(* IEC 61131-3 sources: volt/packages/volt-lsp-iec/test-corpus/pro2193/Device/Plc Logic/Application/09 Misc/Library Manager/L_TT1P_TechnologyModules, 514 files *)

(* ---- _SCAP_TM_BASICMOTIONBASE.dut ---- *)
TYPE _SCAP_TM_BASICMOTIONBASE :
STRUCT
END_STRUCT
END_TYPE

(* ---- _SCAP_TM_BASICMOTIONHIGH.dut ---- *)
TYPE _SCAP_TM_BASICMOTIONHIGH :
STRUCT
END_STRUCT
END_TYPE

(* ---- _SCAP_TM_BASICMOTIONSTATE.dut ---- *)
TYPE _SCAP_TM_BASICMOTIONSTATE :
STRUCT
END_STRUCT
END_TYPE

(* ---- _SCAP_TM_CROSSCUTTERBASE.dut ---- *)
TYPE _SCAP_TM_CROSSCUTTERBASE :
STRUCT
	AP01_XENDOFPROFILEWINDOWSIZE : BOOL;
	AP01_LRENDOFPROFILEWINDOWSIZE : LREAL := 0;
	AP02_XOVERSPEEDUPPERLIMIT : BOOL;
	AP02_LROVERSPEEDUPPERLIMIT : LREAL := 2;
	AP07_XSETOFFSETSLAVE : BOOL;
	AP07_LRSETOFFSETSLAVE : LREAL;
	AP08_XOFFSETSLAVEPAR : BOOL;
	AP08_LROFFSETSLAVEVEL : LREAL;
	AP08_LROFFSETSLAVEACC : LREAL;
	AP08_LROFFSETSLAVEDEC : LREAL;
	AP08_LROFFSETSLAVEJERK : LREAL;
	AP09_XSETVALUEMODE : BOOL;
	AP09_ESETVALUEMODE : L_MC1P_SetValueMode := L_MC1P_SetValueMode.PosVelAcc;
END_STRUCT
END_TYPE

(* ---- _SCAP_TM_CROSSCUTTERHIGH.dut ---- *)
TYPE _SCAP_TM_CROSSCUTTERHIGH :
STRUCT
END_STRUCT
END_TYPE

(* ---- _SCAP_TM_CROSSCUTTERSTATE.dut ---- *)
TYPE _SCAP_TM_CROSSCUTTERSTATE :
STRUCT
	AP03_XTPAXISDELAYCYCLE : BOOL;
	AP03_LRTPAXISDELAYCYCLE : LREAL;
	AP04_XTPAXISCOMPFACTOR : BOOL;
	AP04_LRTPAXISCOMPFACTOR : LREAL;
	AP05_XUPPERCORRPOS : BOOL;
	AP05_LRUPPERCORRPOS : LREAL;
	AP06_XLOWERCORRPOS : BOOL;
	AP06_LRLOWERCORRPOS : LREAL;
	AP10_XCUTTINGANGLESTOPCAM : BOOL;
	AP10_LRCUTTINGANGLESTOPCAM : LREAL := 10;
	AP11_XSETCUTLENGTHINPRODUCT : BOOL;
END_STRUCT
END_TYPE

(* ---- _SCAP_TM_ELECTRICALSHAFTPOSBASE.dut ---- *)
TYPE _SCAP_TM_ELECTRICALSHAFTPOSBASE :
STRUCT
	AP01_XLOADGEARBOXPOSOUT : BOOL;
	AP01_LRLOADGEARBOXPOSOUT : LREAL;
END_STRUCT
END_TYPE

(* ---- _SCAP_TM_ELECTRICALSHAFTPOSHIGH.dut ---- *)
TYPE _SCAP_TM_ELECTRICALSHAFTPOSHIGH :
STRUCT
	AP05_XLOADOFFSETSYNC : BOOL;
	AP05_LRLOADOFFSETSYNC : LREAL;
END_STRUCT
END_TYPE

(* ---- _SCAP_TM_ELECTRICALSHAFTPOSSTATE.dut ---- *)
TYPE _SCAP_TM_ELECTRICALSHAFTPOSSTATE :
STRUCT
	AP02_XLOADTRIMOFFSET : BOOL;
	AP02_LRLOADTRIMOFFSET : LREAL;
END_STRUCT
END_TYPE

(* ---- _SCAP_TM_ELECTRICALSHAFTVELBASE.dut ---- *)
TYPE _SCAP_TM_ELECTRICALSHAFTVELBASE :
STRUCT
	AP01_XCOUPLINGX : BOOL;
	AP01_LRCOUPLINGX : LREAL := 1.0;
	AP02_XCOUPLINGY : BOOL;
	AP02_LRCOUPLINGY : LREAL := 1.0;
END_STRUCT
END_TYPE

(* ---- _SCAP_TM_ELECTRICALSHAFTVELHIGH.dut ---- *)
TYPE _SCAP_TM_ELECTRICALSHAFTVELHIGH :
STRUCT
END_STRUCT
END_TYPE

(* ---- _SCAP_TM_ELECTRICALSHAFTVELSTATE.dut ---- *)
TYPE _SCAP_TM_ELECTRICALSHAFTVELSTATE :
STRUCT
END_STRUCT
END_TYPE

(* ---- _SCAP_TM_FLEXCAMBASE.dut ---- *)
TYPE _SCAP_TM_FLEXCAMBASE :
STRUCT
	AP01_XENDOFPROFILEWINDOWSIZE : BOOL;
	AP01_LRENDOFPROFILEWINDOWSIZE : LREAL := 0;
	AP02_XSETVALUEMODE : BOOL;
	AP02_ESETVALUEMODE : L_MC1P_SetValueMode := L_MC1P_SetValueMode.PosVelAcc;
END_STRUCT
END_TYPE

(* ---- _SCAP_TM_FLEXCAMHIGH.dut ---- *)
TYPE _SCAP_TM_FLEXCAMHIGH :
STRUCT
END_STRUCT
END_TYPE

(* ---- _SCAP_TM_FLEXCAMSTATE.dut ---- *)
TYPE _SCAP_TM_FLEXCAMSTATE :
STRUCT
END_STRUCT
END_TYPE

(* ---- _SCAP_TM_FLYINGSAWBASE.dut ---- *)
TYPE _SCAP_TM_FLYINGSAWBASE :
STRUCT
	AP01_XLOADTOTALCUTTINGLENGTH : BOOL;
	AP01_LRLOADTOTALCUTTINGLENGTH : LREAL;
	AP02_XLOADTARGETPOS : BOOL;
	AP02_LRLOADTARGETPOS : LREAL;
END_STRUCT
END_TYPE

(* ---- _SCAP_TM_FLYINGSAWHIGH.dut ---- *)
TYPE _SCAP_TM_FLYINGSAWHIGH :
STRUCT
	AP02_XLOADTRIMOFFSET : BOOL;
	AP02_LRLOADTRIMOFFSET : LREAL;
END_STRUCT
END_TYPE

(* ---- _SCAP_TM_FLYINGSAWSTATE.dut ---- *)
TYPE _SCAP_TM_FLYINGSAWSTATE :
STRUCT
	AP03_XRANGEOFTOLERANCE : BOOL;
	AP03_LRRANGEOFTOLERANCE : LREAL;
	AP04_XMARKDETECTERRCOMP : BOOL;
	AP04_LRMARKDETECTERRCOMP : LREAL;
	AP05_XTASKCYCLEDELAY : BOOL;
	AP05_BYTASKCYCLEDELAY : BYTE;
END_STRUCT
END_TYPE

(* ---- _SCAP_TM_MOTIONCONTROL.dut ---- *)
TYPE _SCAP_TM_MOTIONCONTROL :
STRUCT
END_STRUCT
END_TYPE

(* ---- _SCAP_TM_PICKANDPLACEBASE.dut ---- *)
TYPE _SCAP_TM_PICKANDPLACEBASE :
STRUCT
	AP01_XCALCPROFILEMOVEPATH : BOOL := TRUE;
END_STRUCT
END_TYPE

(* ---- _SCAP_TM_PICKANDPLACEHIGH.dut ---- *)
TYPE _SCAP_TM_PICKANDPLACEHIGH :
STRUCT
END_STRUCT
END_TYPE

(* ---- _SCAP_TM_PICKANDPLACESTATE.dut ---- *)
TYPE _SCAP_TM_PICKANDPLACESTATE :
STRUCT
	AP02_EBUFFERMODEBLENDING : MC_BUFFER_MODE := MC_BUFFER_MODE.mcBlendingLow;
END_STRUCT
END_TYPE

(* ---- _SCAP_TM_REGISTERCONTROLBASE.dut ---- *)
TYPE _SCAP_TM_REGISTERCONTROLBASE :
STRUCT
	AP03_XTPAXISDELAYCYCLE : BOOL;
	AP03_LRTPAXISDELAYCYCLE : LREAL;
	AP04_XTPAXISCOMPFACTOR : BOOL;
	AP04_LRTPAXISCOMPFACTOR : LREAL;
	AP06_XCORRECTIONONMASTERPOS : BOOL;
	AP07_XLOADSENSORPOS : BOOL;
	AP07_LRLOADSENSORPOS : LREAL;
END_STRUCT
END_TYPE

(* ---- _SCAP_TM_REGISTERCONTROLHIGH.dut ---- *)
TYPE _SCAP_TM_REGISTERCONTROLHIGH :
STRUCT
END_STRUCT
END_TYPE

(* ---- _SCAP_TM_REGISTERCONTROLSTATE.dut ---- *)
TYPE _SCAP_TM_REGISTERCONTROLSTATE :
STRUCT
END_STRUCT
END_TYPE

(* ---- _SCAP_TM_SMARTTRACKBASE.dut ---- *)
TYPE _SCAP_TM_SMARTTRACKBASE :
STRUCT
END_STRUCT
END_TYPE

(* ---- _SCAP_TM_SMARTTRACKHIGH.dut ---- *)
TYPE _SCAP_TM_SMARTTRACKHIGH :
STRUCT
END_STRUCT
END_TYPE

(* ---- _SCAP_TM_SMARTTRACKSTATE.dut ---- *)
TYPE _SCAP_TM_SMARTTRACKSTATE :
STRUCT
	AP_XALLTRACKCORRCAM : BOOL;
	AP_ASCALLTRACKCORRCAM : ARRAY [0..4] OF L_MC2P_XYVA := [STRUCT(eLawOfMotion := L_MC2P_LawOfMotion.Poly5, lrX := 0, lrY := 0, lrYs := 0, lrYss := 0), STRUCT(eLawOfMotion := L_MC2P_LawOfMotion.StraightLine, lrX := 0.179999992251396, lrY := 0.1, lrYs := 1.25000011525118, lrYss := 0), STRUCT(eLawOfMotion := L_MC2P_LawOfMotion.Poly5, lrX := 0.819999933242798, lrY := 0.9, lrYs := 1.25000011525118, lrYss := 0), STRUCT(eLawOfMotion := L_MC2P_LawOfMotion.Poly5, lrX := 1.0, lrY := 1.0, lrYs := 0, lrYss := 0)];
END_STRUCT
END_TYPE

(* ---- _SCAP_TM_STACKERCRANEAXISCONTROLBASE.dut ---- *)
TYPE _SCAP_TM_STACKERCRANEAXISCONTROLBASE :
STRUCT
	AP01_XSETCONTROLLERMODE : BOOL;
	AP01_ECONTROLMODE : L_MC1P_ControlModeSet;
	AP03_XOSCCOMPPOSSCALED : BOOL;
	AP03_LROSCCOMPPOSSCALED : LREAL;
	AP04_XOSCCOMPLOADSCALED : BOOL;
	AP04_LROSCCOMPLOADSCALED : LREAL;
	AP05_EOSCCOMPEXECUTIONINDEX : WORD := 1;
	AP06_XOSCCOMPIGNOREFILTERONSTOP : BOOL := FALSE;
	AP07_XOSCCOMPMANIPULATETROQUE : BOOL := FALSE;
	AP08_XOSCCOMPAMPRATIO : BOOL;
	AP08_LROSCCOMPAMPRATIO : LREAL;
	AP09_XOSCCOMPEIGENFREQ : BOOL;
	AP09_LROSCCOMPEIGENFREQ : LREAL;
	AP10_XUPDATEEIGENFREQ : BOOL;
	AP11_XUPDATEAMPRATIO : BOOL;
	AP12_XWAITFORBRAKERELEASED : BOOL;
	AP13_XBRAKETESTMODE : BOOL;
	AP13_EBRAKETESTMODE : L_MC1P_BrakeTestMode;
	AP14_XBRAKETESTDIRECTION : BOOL;
	AP14_EBRAKETESTDIRECTION : MC_DIRECTION;
	AP18_XBRAKEGRINDINMODE : BOOL;
	AP18_EBRAKEGRINDINMODE : L_MC1P_GrindInMode;
	AP20_XFILTTIMEACTTORQUE : BOOL;
	AP20_LRFILTTIMEACTTORQUE : LREAL := 0.02;
END_STRUCT
END_TYPE

(* ---- _SCAP_TM_STACKERCRANEHEADCONTROLBASE.dut ---- *)
TYPE _SCAP_TM_STACKERCRANEHEADCONTROLBASE :
STRUCT
END_STRUCT
END_TYPE

(* ---- _SCAP_TM_TABLEPOSITIONINGBASE.dut ---- *)
TYPE _SCAP_TM_TABLEPOSITIONINGBASE :
STRUCT
END_STRUCT
END_TYPE

(* ---- _SCAP_TM_WINDER.dut ---- *)
TYPE _SCAP_TM_WINDER :
STRUCT
	AP09_XSETVELOFFSET : BOOL;
	AP09_LRSETVELOFFSET : LREAL;
	AP10_XSETTRQOFFSET : BOOL;
	AP10_LRSETTRQOFFSET : LREAL;
	AP11_XSETVELOFFSETDIAMCACL : BOOL;
	AP11_LRSETVELOFFSETDIAMCACL : LREAL;
	AP12_XSETSPEEDPOINTDIAMCALC : BOOL;
	AP12_LRSETSPEEDPOINTDIAMCALC : LREAL;
END_STRUCT
END_TYPE

(* ---- _SCAP_TM_WINDERDANCERCTRLBASE.dut ---- *)
TYPE _SCAP_TM_WINDERDANCERCTRLBASE :
STRUCT
	AP01_XSETSPEEDPOINT : BOOL;
	AP01_LRSETSPEEDPOINT : LREAL;
	AP03_XSETDANCERCTRLOUTGAIN : BOOL;
	AP03_LRSETDANCERCTRLOUTGAIN : LREAL;
	AP04_XSETDANCERCTRLOUTRESETTIME : BOOL;
	AP04_LRSETDANCERCTRLOUTRESETTIME : LREAL;
	AP05_XSETDANCERCTRLOUTRATETIME : BOOL;
	AP05_LRSETDANCERCTRLOUTRATETIME : LREAL;
END_STRUCT
END_TYPE

(* ---- _SCAP_TM_WINDERDANCERCTRLHIGH.dut ---- *)
TYPE _SCAP_TM_WINDERDANCERCTRLHIGH :
STRUCT
END_STRUCT
END_TYPE

(* ---- _SCAP_TM_WINDERDANCERCTRLSTATE.dut ---- *)
TYPE _SCAP_TM_WINDERDANCERCTRLSTATE :
STRUCT
	AP02_XSETTRQPOINT : BOOL;
	AP02_LRSETTRQPOINT : LREAL;
END_STRUCT
END_TYPE

(* ---- _SCAP_TM_WINDERTENSIONCTRLBASE.dut ---- *)
TYPE _SCAP_TM_WINDERTENSIONCTRLBASE :
STRUCT
	AP1_XSETACCCOMPTRQ : BOOL;
	AP1_LRSETACCCOMPTRQ : LREAL;
	AP02_XSETTRQPOINT : BOOL;
	AP02_LRSETTRQPOINT : LREAL;
	AP3_XSETUPPERSPEEDLIMIT : BOOL;
	AP3_LRSETUPPERSPEEDLIMIT : LREAL;
	AP4_XSETLOWERSPEEDLIMIT : BOOL;
	AP4_LRSETLOWERSPEEDLIMIT : LREAL;
END_STRUCT
END_TYPE

(* ---- _SCAP_TM_WINDERTENSIONCTRLHIGH.dut ---- *)
TYPE _SCAP_TM_WINDERTENSIONCTRLHIGH :
STRUCT
END_STRUCT
END_TYPE

(* ---- _SCAP_TM_WINDERTENSIONCTRLSTATE.dut ---- *)
TYPE _SCAP_TM_WINDERTENSIONCTRLSTATE :
STRUCT
	AP05_XSETTENSIONCTRLOUTGAIN : BOOL;
	AP05_LRSETTENSIONCTRLOUTGAIN : LREAL;
	AP06_XSETTENSIONCTRLOUTRESETTIME : BOOL;
	AP06_LRSETTENSIONCTRLOUTRESETTIME : LREAL;
	AP07_XSETTENSIONCTRLOUTRATETIME : BOOL;
	AP07_LRSETTENSIONCTRLOUTRATETIME : LREAL;
	AP08_XSETFRICCOMPREELSPEED : BOOL;
	AP08_LRSETFRICCOMPREELSPEED : LREAL;
END_STRUCT
END_TYPE

(* ---- _SCPAR_TM_BASE.dut ---- *)
TYPE _SCPAR_TM_BASE :
STRUCT
END_STRUCT
END_TYPE

(* ---- _SCPAR_TM_BASICMOTIONBASE.dut ---- *)
TYPE _SCPAR_TM_BASICMOTIONBASE :
STRUCT
	LRVEL : LREAL := 50;
	LRACC : LREAL := 100;
	LRDEC : LREAL := 100;
	EDIRECTION : MC_DIRECTION := MC_DIRECTION.mcPositiveDirection;
	XCONTINUOUSUPDATE : BOOL;
END_STRUCT
END_TYPE

(* ---- _SCPAR_TM_BASICMOTIONHIGH.dut ---- *)
TYPE _SCPAR_TM_BASICMOTIONHIGH :
STRUCT
END_STRUCT
END_TYPE

(* ---- _SCPAR_TM_BASICMOTIONSTATE.dut ---- *)
TYPE _SCPAR_TM_BASICMOTIONSTATE :
STRUCT
END_STRUCT
END_TYPE

(* ---- _SCPAR_TM_CROSSCUTTERBASE.dut ---- *)
TYPE _SCPAR_TM_CROSSCUTTERBASE :
STRUCT
	ETRIMMODE : L_TT1P_TrimMode := L_TT1P_TrimMode.position;
	LRTRIMDIST : LREAL := 3;
	LROFFSETTRIMVEL : LREAL := 10;
	LROFFSETTRIMACC : LREAL := 100;
	LROFFSETTRIMDEC : LREAL := 100;
	EPOSITIONINGDIRECTION : MC_DIRECTION := MC_DIRECTION.mcPositiveDirection;
	LRPOSITIONINGVEL : LREAL := 10;
	LRPOSITIONINGACC : LREAL := 100;
	LRPOSITIONINGDEC : LREAL := 100;
	ESYNCMODE : L_TT1P_SyncModeCrossCutter;
	LRMASTERSYNCINDIST : LREAL := 0;
	LRMASTERSYNCOUTDIST : LREAL := 0;
	LRSYNCOUTINSTANTDEC : LREAL := 1000;
	XMASTERABSOLUTE : BOOL := TRUE;
	LRSTARTXPOSRELATIVE : LREAL := 0;
	BYSTARTTOOLNO : BYTE := 0;
	BYNUMOFTOOLS : BYTE := 1;
	LRCUTTINGANGLE : LREAL := 10;
	LRCROSSCUTTERCIRCUMFERENCE : LREAL := 75.55555;
	LRSCALINGMASTER : LREAL := 1;
	XCALCCAMBOUNDS : BOOL := FALSE;
	LRMASTERMAXVEL : LREAL := 100;
	LRMASTERMAXACC : LREAL := 1000;
	EPROFILETYPE : L_MC2P_LawOfMotion := L_MC2P_LawOfMotion.Poly5;
END_STRUCT
END_TYPE

(* ---- _SCPAR_TM_CROSSCUTTERBASEEXTENSION.dut ---- *)
TYPE _SCPAR_TM_CROSSCUTTERBASEEXTENSION :
STRUCT
	ECUTTINGMODE : L_TT1P_CuttingModeBase := L_TT1P_CuttingModeBase.cut_length;
END_STRUCT
END_TYPE

(* ---- _SCPAR_TM_CROSSCUTTERHIGH.dut ---- *)
TYPE _SCPAR_TM_CROSSCUTTERHIGH :
STRUCT
END_STRUCT
END_TYPE

(* ---- _SCPAR_TM_CROSSCUTTERSTATE.dut ---- *)
TYPE _SCPAR_TM_CROSSCUTTERSTATE :
STRUCT
	ECUTTINGMODE : L_TT1P_CuttingModeState;
	ALRCUTLENGTHINPRODUCT : ARRAY [1..10] OF LREAL;
	LRMINPRODUCTLENGTH : LREAL := 50;
	LRTRQCTRLGAIN : LREAL := 0;
	LRTRQCTRLRATETIME : LREAL := 0;
	LRMINERTIA : LREAL := 0;
	LRSENSORTOOLDIST : LREAL := 0.0;
	XMARKCORRECTION : BOOL := TRUE;
	LRMARKWINDOWSIZE : LREAL := 20;
	LRSETOFFSETMARKWINDOW : LREAL := 0.0;
	ETPMODE : L_TT1P_TpMode := L_TT1P_TpMode.TpFromMaster;
	LRCYCLELENGTHEXTENCODER : LREAL := 360;
	LRMAXCORRPOS : LREAL := 30.0;
	LRMAXCORRNEG : LREAL := -30.0;
	LRGEARFACTORCORRGAIN : LREAL := 0.1;
	LRMAXGEARFACTORCORR : LREAL := 10;
	DWMAXMISSEDMARKS : DWORD := 5;
END_STRUCT
END_TYPE

(* ---- _SCPAR_TM_ELECTRICALSHAFTPOSBASE.dut ---- *)
TYPE _SCPAR_TM_ELECTRICALSHAFTPOSBASE :
STRUCT
	DWNUMERATOR : DWORD := 1;
	DWDENOMINATOR : DWORD := 1;
	XLOADSYNCPOS : BOOL;
END_STRUCT
END_TYPE

(* ---- _SCPAR_TM_ELECTRICALSHAFTPOSHIGH.dut ---- *)
TYPE _SCPAR_TM_ELECTRICALSHAFTPOSHIGH :
STRUCT
	EOFFSETMASTERDIRECTION : L_TT1P_Direction;
	EOFFSETMASTERPROFILETYPE : L_TT1P_ProfileType := L_TT1P_ProfileType.poly_5th_order;
	LROFFSETMASTERVELPOS : LREAL := 100.0;
	LROFFSETMASTERVELNEG : LREAL := 100.0;
	LROFFSETMASTERACCDEC : LREAL := 1000.0;
	XLOADOFFSETMASTER : BOOL;
	EOFFSETSLAVEDIRECTION : L_TT1P_Direction := L_TT1P_Direction.DirectionMaster;
	EOFFSETSLAVEPROFILETYPE : L_TT1P_ProfileType := 2;
	LROFFSETSLAVEVELPOS : LREAL := 100.0;
	LROFFSETSLAVEVELNEG : LREAL := 100.0;
	LROFFSETSLAVEACCDEC : LREAL := 1000.0;
	XLOADOFFSETSLAVE : BOOL;
	ESYNCSLAVEDIRECTION : L_TT1P_SyncDirectionElectricalShaftPos := L_TT1P_SyncDirectionElectricalShaftPos.mcShortestWay;
	ESYNCMODE : L_TT1P_SyncModeElectricalShaftPos := L_TT1P_SyncModeElectricalShaftPos.Ramp_Dist;
	LRSYNCINTIME : LREAL := 5;
	LRSYNCOUTTIME : LREAL := 5;
	LRSYNCVEL : LREAL := 100;
	LRSYNCACC : LREAL := 1000.0;
	LRSYNCDEC : LREAL := 1000.0;
	LRSYNCJERK : LREAL := 1000000.0;
	LRSYNCOUTINSTANTDEC : LREAL := 10000;
END_STRUCT
END_TYPE

(* ---- _SCPAR_TM_ELECTRICALSHAFTPOSSTATE.dut ---- *)
TYPE _SCPAR_TM_ELECTRICALSHAFTPOSSTATE :
STRUCT
	LRTRIMACC : LREAL := 100;
	LRTRIMDEC : LREAL := 100;
	LRTRIMVEL : LREAL := 50;
	LRSLAVESYNCINDIST : LREAL := 90.0;
	LRSLAVESYNCOUTDIST : LREAL := 90.0;
	LRSLAVESYNCOUTPOS : LREAL := 0.0;
END_STRUCT
END_TYPE

(* ---- _SCPAR_TM_ELECTRICALSHAFTVELBASE.dut ---- *)
TYPE _SCPAR_TM_ELECTRICALSHAFTVELBASE :
STRUCT
	DWCOUPLINGMODE : DWORD := 1;
	LRCOUPLINGX : LREAL := 1.0;
	LRCOUPLINGY : LREAL := 1.0;
END_STRUCT
END_TYPE

(* ---- _SCPAR_TM_ELECTRICALSHAFTVELHIGH.dut ---- *)
TYPE _SCPAR_TM_ELECTRICALSHAFTVELHIGH :
STRUCT
	LROFFSETACC : LREAL := 100.0;
	LROFFSETDEC : LREAL := 100.0;
	LROFFSETJERK : LREAL := 10000;
END_STRUCT
END_TYPE

(* ---- _SCPAR_TM_ELECTRICALSHAFTVELSTATE.dut ---- *)
TYPE _SCPAR_TM_ELECTRICALSHAFTVELSTATE :
STRUCT
	LRTRIMACC : LREAL := 100;
	LRTRIMDEC : LREAL := 100;
	LRTRIMVEL : LREAL := 50;
	LRSYNCOUTACC : LREAL := 100.0;
	LRSYNCINACC : LREAL := 100.0;
	LRSYNCJERK : LREAL := 10000;
END_STRUCT
END_TYPE

(* ---- _SCPAR_TM_FLEXCAMBASE.dut ---- *)
TYPE _SCPAR_TM_FLEXCAMBASE :
STRUCT
	ESYNCMODE : L_TT1P_SyncMode := L_TT1P_SyncMode.absolute;
	ESYNCDIRECTION : L_TT1P_SyncDirection := L_TT1P_SyncDirection.mcCurrentDirection;
	LRMASTERSYNCINDIST : LREAL := 100;
	LRMASTERSYNCINPOS : LREAL := 0;
	LRMASTERSYNCOUTDIST : LREAL := 100;
	LRSLAVESYNCOUTPOS : LREAL := 0;
	LRSYNCINTIME : LREAL := 5;
	LRSYNCOUTTIME : LREAL := 5;
	LRSYNCOUTINSTANTDEC : LREAL := 10000;
	LRSYNCVEL : LREAL := 100;
	LRSYNCACC : LREAL := 1000.0;
	LRSYNCDEC : LREAL := 1000.0;
	LRSYNCJERK : LREAL := 1000000.0;
	XCAMCYCLIC : BOOL := TRUE;
	XMASTERABSOLUTE : BOOL := TRUE;
	XSLAVEABSOLUTE : BOOL := TRUE;
	EOFFSETMODEMASTER : L_TT1P_OffsetMode := ANY_TO_WORD(L_TT1P_OffsetMode.x_zero);
	EOFFSETMODESLAVE : L_TT1P_OffsetModeSlave := ANY_TO_WORD(L_TT1P_OffsetMode.x_zero);
	LROFFSETSCALINGMASTERVEL : LREAL := 100.0;
	LROFFSETSCALINGMASTERACC : LREAL := 1000.0;
	LROFFSETSCALINGMASTERDEC : LREAL := 1000.0;
	ESCALINGMODEMASTER : L_TT1P_ScalingMode := L_TT1P_ScalingMode.x_zero;
	ESCALINGMODESLAVE : L_TT1P_ScalingMode := L_TT1P_ScalingMode.x_zero;
	LROFFSETSCALINGSLAVEVEL : LREAL := 100.0;
	LROFFSETSCALINGSLAVEACC : LREAL := 1000.0;
	LROFFSETSCALINGSLAVEDEC : LREAL := 1000.0;
	XCALCCAMBOUNDS : BOOL;
	LRMASTERMAXVEL : LREAL := 100;
	LRMASTERMAXACC : LREAL := 1000;
END_STRUCT
END_TYPE

(* ---- _SCPAR_TM_FLEXCAMHIGH.dut ---- *)
TYPE _SCPAR_TM_FLEXCAMHIGH :
STRUCT
END_STRUCT
END_TYPE

(* ---- _SCPAR_TM_FLEXCAMSTATE.dut ---- *)
TYPE _SCPAR_TM_FLEXCAMSTATE :
STRUCT
	EPOSCTRLDIRECTION : L_TT1P_Direction := L_TT1P_Direction.both;
	ECAMSEQUENCEMODE : L_TT1P_CamSequenceMode := L_TT1P_CamSequenceMode.CyclicCam1;
END_STRUCT
END_TYPE

(* ---- _SCPAR_TM_FLYINGSAWBASE.dut ---- *)
TYPE _SCPAR_TM_FLYINGSAWBASE :
STRUCT
	LRSYNCVEL : LREAL := 3600;
	LRSYNCACC : LREAL := 10000;
	LRSYNCDEC : LREAL := 10000;
	LRPOSVEL : LREAL := 3600;
	LRPOSACC : LREAL := 10000;
	LRPOSDEC : LREAL := 10000;
	LRSETMATERIALPOS : LREAL := 0;
	LRUPPERLIMIT : LREAL := 1000;
	LRLOWERLIMIT : LREAL := 0;
	LRGAP : LREAL;
	LRBLADEWIDTH : LREAL := 0;
	XSYNCFLYINGSAW : BOOL := FALSE;
END_STRUCT
END_TYPE

(* ---- _SCPAR_TM_FLYINGSAWHIGH.dut ---- *)
TYPE _SCPAR_TM_FLYINGSAWHIGH :
STRUCT
	EOFFSETSLAVEDIRECTION : L_TT1P_Direction := L_TT1P_Direction.DirectionMaster;
	EOFFSETSLAVEPROFILETYPE : L_TT1P_ProfileType := 2;
	LROFFSETSLAVEVELPOS : LREAL := 10000.0;
	LROFFSETSLAVEVELNEG : LREAL := 10000.0;
	LROFFSETSLAVEACCDEC : LREAL := 10000.0;
	XLOADOFFSETSLAVE : BOOL;
END_STRUCT
END_TYPE

(* ---- _SCPAR_TM_FLYINGSAWSTATE.dut ---- *)
TYPE _SCPAR_TM_FLYINGSAWSTATE :
STRUCT
	XPARKPOS : BOOL := FALSE;
	LRPARKPOSITION : LREAL := 0;
	LRMARKSENSORPOS : LREAL;
	EMODEFLYINGSAW : L_TT1P_eModesFlyingSaw;
	XPOSINWINDOW : BOOL;
	LRPOSINWINDOW : LREAL;
	LRTIMEPOSINWINDOW : LREAL := 50;
END_STRUCT
END_TYPE

(* ---- _SCPAR_TM_MOTIONCONTROL.dut ---- *)
TYPE _SCPAR_TM_MOTIONCONTROL :
STRUCT
	LRSTOPDEC : LREAL := 10000;
	LRSTOPJERK : LREAL := 100000;
	LRHALTDEC : LREAL := 3600;
	LRJERK : LREAL := 100000;
END_STRUCT
END_TYPE

(* ---- _SCPAR_TM_MOTIONCONTROLAGBC.dut ---- *)
TYPE _SCPAR_TM_MOTIONCONTROLAGBC :
STRUCT
	LRPATHSTOPDEC : LREAL := 10000;
	LRPATHSTOPJERK : LREAL := 100000;
	LRPATHHALTDEC : LREAL := 100;
	LRPATHJERK : LREAL := 100000;
	ALRSTOPDEC : ARRAY [1..18] OF LREAL := [18(10000)];
	ALRSTOPJERK : ARRAY [1..18] OF LREAL := [18(100000)];
END_STRUCT
END_TYPE

(* ---- _SCPAR_TM_MOTIONCONTROLBASE.dut ---- *)
TYPE _SCPAR_TM_MOTIONCONTROLBASE :
STRUCT
	LRJOGJERK : LREAL := 10000;
	LRJOGVEL : LREAL := 10;
	LRJOGACC : LREAL := 100;
	LRJOGDEC : LREAL := 100;
END_STRUCT
END_TYPE

(* ---- _SCPAR_TM_MOTIONCONTROLSTATE.dut ---- *)
TYPE _SCPAR_TM_MOTIONCONTROLSTATE :
STRUCT
	LRHOMEPOSITION : LREAL := 0;
	XUSEHOMEEXTPARAMETER : BOOL := FALSE;
	SCHOMEEXTPARAMETER : L_MC1P_HomeParameter := STRUCT(eHomeMode := L_MC1P_HomeMode.SetPositionDirect);
	SCHOMEEXTTP : MC_TRIGGER_REF;
END_STRUCT
END_TYPE

(* ---- _SCPAR_TM_PICKANDPLACEBASE.dut ---- *)
TYPE _SCPAR_TM_PICKANDPLACEBASE :
STRUCT
	LRCARTESIANJOGJERK : LREAL := 10000;
	LRCARTESIANJOGVEL : LREAL := 10;
	LRCARTESIANJOGACC : LREAL := 100;
	LRCARTESIANJOGDEC : LREAL := 100;
	LRORIENTATIONJOGJERK : LREAL := 10000;
	LRORIENTATIONJOGVEL : LREAL := 10;
	LRORIENTATIONJOGACC : LREAL := 100;
	LRORIENTATIONJOGDEC : LREAL := 100;
	LRREALAXISJOGJERK : LREAL := 10000;
	LRREALAXISJOGVEL : LREAL := 10;
	LRREALAXISJOGACC : LREAL := 100;
	LRREALAXISJOGDEC : LREAL := 100;
	ALRHOMEPOSITION : ARRAY [1..12] OF LREAL;
	AEHOMINGORDER : ARRAY [1..12] OF L_MC4P_HomingOrder;
	XUSEHOMEEXTPARAMETER : BOOL := FALSE;
	ASCHOMEEXTTP : ARRAY [1..12] OF MC_TRIGGER_REF;
	ASCHOMEEXTPARAMETER : ARRAY [1..12] OF L_MC1P_HomeParameter := [STRUCT(eHomeMode := L_MC1P_HomeMode.SetPositionDirect), STRUCT(eHomeMode := L_MC1P_HomeMode.SetPositionDirect), STRUCT(eHomeMode := L_MC1P_HomeMode.SetPositionDirect), STRUCT(eHomeMode := L_MC1P_HomeMode.SetPositionDirect), STRUCT(eHomeMode := L_MC1P_HomeMode.SetPositionDirect), STRUCT(eHomeMode := L_MC1P_HomeMode.SetPositionDirect), STRUCT(eHomeMode := L_MC1P_HomeMode.SetPositionDirect), STRUCT(eHomeMode := L_MC1P_HomeMode.SetPositionDirect), STRUCT(eHomeMode := L_MC1P_HomeMode.SetPositionDirect), STRUCT(eHomeMode := L_MC1P_HomeMode.SetPositionDirect), STRUCT(eHomeMode := L_MC1P_HomeMode.SetPositionDirect), STRUCT(eHomeMode := L_MC1P_HomeMode.SetPositionDirect)];
	LRXMAXVEL : LREAL := 10;
	LRYMAXVEL : LREAL := 10;
	LRZMAXVEL : LREAL := 10;
	LRAMAXVEL : LREAL := 10;
	LRBMAXVEL : LREAL := 10;
	LRCMAXVEL : LREAL := 10;
	LRAUX1MAXVEL : LREAL := 10;
	LRXMAXACCDEC : LREAL := 100;
	LRYMAXACCDEC : LREAL := 100;
	LRZMAXACCDEC : LREAL := 100;
	LRAMAXACCDEC : LREAL := 100;
	LRBMAXACCDEC : LREAL := 100;
	LRCMAXACCDEC : LREAL := 100;
	LRAUX1MAXACCDEC : LREAL := 100;
	LRXMAXJERK : LREAL := 10000;
	LRYMAXJERK : LREAL := 10000;
	LRZMAXJERK : LREAL := 10000;
	LRAMAXJERK : LREAL := 10000;
	LRBMAXJERK : LREAL := 10000;
	LRCMAXJERK : LREAL := 10000;
	LRAUX1MAXJERK : LREAL := 10000;
	LRGRIPPERCLOSINGTIME : LREAL;
	XPOSINWINDOW : BOOL;
	LRPOSINWINDOW : LREAL := 0.5;
	LRTIMEPOSINWINDOW : LREAL := 50;
END_STRUCT
END_TYPE

(* ---- _SCPAR_TM_PICKANDPLACEBASEEXTENSION.dut ---- *)
TYPE _SCPAR_TM_PICKANDPLACEBASEEXTENSION :
STRUCT
	ETARGETCOORDSYSTEM : L_MC4P_CoordSystem := 0;
	LRXTARGETPOS : LREAL;
	LRYTARGETPOS : LREAL;
	LRZTARGETPOS : LREAL;
	LRATARGETPOS : LREAL := 180;
	LRBTARGETPOS : LREAL;
	LRCTARGETPOS : LREAL;
	LRAUX1TARGETPOS : LREAL;
	LRZSTARTDIST : LREAL;
	LRZTARGETDIST : LREAL;
	LRBLENDINGRADIUS : LREAL;
	LRPATHVEL : LREAL := 10;
	LRPATHACC : LREAL := 100;
	LRPATHDEC : LREAL := 100;
END_STRUCT
END_TYPE

(* ---- _SCPAR_TM_PICKANDPLACEHIGH.dut ---- *)
TYPE _SCPAR_TM_PICKANDPLACEHIGH :
STRUCT
END_STRUCT
END_TYPE

(* ---- _SCPAR_TM_PICKANDPLACESTATE.dut ---- *)
TYPE _SCPAR_TM_PICKANDPLACESTATE :
STRUCT
	XSINGLESTEP : BOOL := FALSE;
	ASCPROFILEPAR : ARRAY [1..10] OF L_TT1P_scProfilePar;
END_STRUCT
END_TYPE

(* ---- _SCPAR_TM_REGISTERCONTROLBASE.dut ---- *)
TYPE _SCPAR_TM_REGISTERCONTROLBASE :
STRUCT
	LRSENSORTOOLDIST : LREAL := 0.0;
	XMARKCORRECTION : BOOL := TRUE;
	LRMARKDIST : LREAL := 360.0;
	LRCYCLELENGTHEXTENCODER : LREAL := 360;
	ETPMODE : L_TT1P_TpMode := L_TT1P_TpMode.TpFromMaster;
	LRMAXCORRPOS : LREAL := 30.0;
	LRMAXCORRNEG : LREAL := -30.0;
	ESOURCEFORCORRWINDOW : L_TT1P_SourceForCorrWindow := L_TT1P_SourceForCorrWindow.Slave;
	LRUPPERCORRPOS : LREAL := 180.0;
	LRLOWERCORRPOS : LREAL := 90.0;
	LRTRIMDIST : LREAL := 1;
	ETRIMMODE : L_TT1P_TrimMode := 0;
END_STRUCT
END_TYPE

(* ---- _SCPAR_TM_REGISTERCONTROLHIGH.dut ---- *)
TYPE _SCPAR_TM_REGISTERCONTROLHIGH :
STRUCT
END_STRUCT
END_TYPE

(* ---- _SCPAR_TM_REGISTERCONTROLSTATE.dut ---- *)
TYPE _SCPAR_TM_REGISTERCONTROLSTATE :
STRUCT
	LRMARKWINDOWSIZE : LREAL := 90.0;
	LRSETOFFSETMARKWINDOW : LREAL := 0.0;
	LRGEARFACTORCORRGAIN : LREAL := 0.1;
	LRMAXGEARFACTORCORR : LREAL := 10;
	DWMAXNUMBERVIRTUALMARKS : DWORD := 5;
END_STRUCT
END_TYPE

(* ---- _SCPAR_TM_SMARTTRACKBASE.dut ---- *)
TYPE _SCPAR_TM_SMARTTRACKBASE :
STRUCT
	LRSYNCINACC : LREAL := 100;
	LRSYNCOUTACC : LREAL := 100;
	LRSYNCJERK : LREAL := 10000;
	XDISABLECORRECTION : BOOL;
	XPITCHCHECK : BOOL := TRUE;
	ETPMODE : L_TT1P_TpMode;
	LRPRODUCTTARGET : LREAL := 0;
	BYNUMOFPRODUCTTARGETS : BYTE := 1;
	LRCORRDISTRIBRUTIONSCALED : LREAL := 0.5;
	LRVELFACTORSCALED : LREAL := 1;
	LRMAXCORRPOS : LREAL := 100;
	LRMAXCORRNEG : LREAL := 100;
	LRCORRDIST : LREAL := 300;
	LRDEBOUNCINGWINDOWEDGERISE : LREAL := 10;
	LRDEBOUNCINGWINDOWEDGEFALL : LREAL := 0;
END_STRUCT
END_TYPE

(* ---- _SCPAR_TM_SMARTTRACKHIGH.dut ---- *)
TYPE _SCPAR_TM_SMARTTRACKHIGH :
STRUCT
END_STRUCT
END_TYPE

(* ---- _SCPAR_TM_SMARTTRACKSTATE.dut ---- *)
TYPE _SCPAR_TM_SMARTTRACKSTATE :
STRUCT
	LRSMARTTRACKLENGTH : LREAL := 300;
	LRSENSORPOSITION : LREAL := 100;
	LRPRODUCTHANDOVERDIST : LREAL := 100;
	XALLTRACKCORRECTION : BOOL := FALSE;
	LRALLTRACKSYNCDIST : LREAL := 50;
END_STRUCT
END_TYPE

(* ---- _SCPAR_TM_STACKERCRANEAXISCONTROLBASE.dut ---- *)
TYPE _SCPAR_TM_STACKERCRANEAXISCONTROLBASE :
STRUCT
	EREGULATORONMODE : L_TT1P_RegulatorOnMode := 0;
	LRDISABLEAFTERTIME : LREAL := 60;
	SCMINLIMITS : L_TT1P_XYLimits;
	SCBUFFERDATA : L_TT1P_XYBufferData;
	XBUFFERRANGE : BOOL;
	LRMAINTENANCEVEL : LREAL := 10;
	LRMAINTENANCEACC : LREAL := 100;
	LRMAINTENANCEDEC : LREAL := 100;
	LRMAINTENANCEJERK : LREAL := 10000;
	EOSCCOMPMODE : L_CT1P.L_CT1P_OscCompMode := 0;
	ASCOSCCOMPDATA : ARRAY [1..8] OF L_TT1P_OscillationCompensationData;
	LRBRAKETESTMOTORTRQ : LREAL;
	LRBRAKETESTRAMPTIME : LREAL;
	LRBRAKETESTHOLDTIME : LREAL;
	LRBRAKETESTPOSTHRESHOLD : LREAL;
	WBRAKEGRINDINCYCLES : WORD;
	EBRAKEGRINDMODE : L_MC1P_GrindInMode;
	LRBRAKEGRINDINMOTORSPEED : LREAL;
	LRBRAKEGRINDINRAMPTIME : LREAL;
	LRBRAKEGRINDINONTIME : LREAL;
	LRBRAKEGRINDINOFFTIME : LREAL;
	EBRAKEGRINDINADDITIONALLIMITS : L_MC1P_AdditionalLimits := L_MC1P_AdditionalLimits.NotActive;
	LRBRAKEGRINDINPOSLIMIT1 : LREAL;
	LRBRAKEGRINDINPOSLIMIT2 : LREAL;
	XBRAKEGRINDINFINISHINSTARTPOS : BOOL;
	XBRAKEEXTERNALFAN : BOOL;
END_STRUCT
END_TYPE

(* ---- _SCPAR_TM_STACKERCRANEHEADCONTROLBASE.dut ---- *)
TYPE _SCPAR_TM_STACKERCRANEHEADCONTROLBASE :
STRUCT
	EXYMODE : L_TT1P_XYMode;
	SCXPROFILE : L_TT1P_MoveAbsProfileData;
	SCYPROFILE : L_TT1P_MoveAbsProfileData;
END_STRUCT
END_TYPE

(* ---- _SCPAR_TM_TABLEPOSITIONINGBASE.dut ---- *)
TYPE _SCPAR_TM_TABLEPOSITIONINGBASE :
STRUCT
	ETPMODE : L_TT1P_TpModeSingleAxis;
	LRCYCLELENGTHEXTENCODER : LREAL := 360;
	SCPROFILES : L_TT1P_Profiles;
	XCONTINUOUSUPDATE : BOOL := FALSE;
	XABSOLUTEMODULOCYCLE : BOOL := FALSE;
	XLOADTORQUELIMITS : BOOL := FALSE;
END_STRUCT
END_TYPE

(* ---- _SCPAR_TM_TABLEPOSITIONINGHIGH.dut ---- *)
TYPE _SCPAR_TM_TABLEPOSITIONINGHIGH :
STRUCT
END_STRUCT
END_TYPE

(* ---- _SCPAR_TM_TABLEPOSITIONINGSTATE.dut ---- *)
TYPE _SCPAR_TM_TABLEPOSITIONINGSTATE :
STRUCT
END_STRUCT
END_TYPE

(* ---- _SCPAR_TM_VIRTUALMASTERBASE.dut ---- *)
TYPE _SCPAR_TM_VIRTUALMASTERBASE :
STRUCT
	LRACC : LREAL := 100;
	LRDEC : LREAL := 100;
	EDIRECTION : MC_DIRECTION := MC_DIRECTION.mcPositiveDirection;
END_STRUCT
END_TYPE

(* ---- _SCPAR_TM_VIRTUALMASTERHIGH.dut ---- *)
TYPE _SCPAR_TM_VIRTUALMASTERHIGH :
STRUCT
	ESYNCMODE : L_TT1P_SyncModeVirtualMaster := L_TT1P_SyncModeVirtualMaster.Ramp_Dist;
	ESYNCSLAVEDIRECTION : L_TT1P_SyncDirectionVirtualMaster := L_TT1P_SyncDirectionVirtualMaster.mcShortestWay;
	LRMASTERSYNCINDIST : LREAL := 90;
	LRSYNCINTIME : LREAL := 5;
	LRSYNCVEL : LREAL := 100;
	LRSYNCACC : LREAL := 1000.0;
	LRSYNCDEC : LREAL := 1000.0;
	LRSYNCJERK : LREAL := 1000000.0;
END_STRUCT
END_TYPE

(* ---- _SCPAR_TM_VIRTUALMASTERSTATE.dut ---- *)
TYPE _SCPAR_TM_VIRTUALMASTERSTATE :
STRUCT
END_STRUCT
END_TYPE

(* ---- _SCPAR_TM_VIRTUALMASTERSTATEEXTENSION.dut ---- *)
TYPE _SCPAR_TM_VIRTUALMASTERSTATEEXTENSION :
STRUCT
	LRMASTERACCDEC : LREAL := 100;
END_STRUCT
END_TYPE

(* ---- _SCPAR_TM_WINDER.dut ---- *)
TYPE _SCPAR_TM_WINDER :
STRUCT
	LRLINEJERK : LREAL := 10000;
	LRJOGLINEACC : LREAL := 100;
	LRJOGLINEDEC : LREAL := 100;
	LRJOGLINEVEL : LREAL := 10;
	LRTRIMLINEACC : LREAL := 100;
	LRTRIMLINEDEC : LREAL := 100;
	LRTRIMLINEVEL : LREAL := 10;
	LRSYNCLINEACC : LREAL := 100;
	LRSYNCLINEDEC : LREAL := 100;
	LRWEBBREAKWINDOW : LREAL := 0.1;
	LRMAXDIAM : LREAL := 180;
	LRMINDIAM : LREAL := 50;
	RFILTTIMEDIAM : REAL := 0.05;
	LRDIAMCALCREGULARDIST : LREAL := 1;
	LRDIAMCALCREDUCEDDIST : LREAL := 0.1;
	ALRADAPTDIAMX : ARRAY [1..9] OF LREAL := [0, 100, 200, 300, 400, 500, 600, 700, 800];
	ALRADAPTDIAMY : ARRAY [1..9] OF LREAL := [0, 100, 200, 300, 400, 500, 600, 700, 800];
	LRTENSCURVECTRLSCALED : LREAL := 0;
	LRTENSCURVESTARTDIAMSCALED : LREAL := 0;
	LRLINEVELREF : LREAL := 1000;
	LRMINLINEVEL : LREAL := 1;
	RFILTTIMEMATERIALCOUNTER : REAL := 0.0;
	LRSETMATERIALPOS : LREAL;
	LRMAXWNDSPD : LREAL := 100;
END_STRUCT
END_TYPE

(* ---- _SCPAR_TM_WINDERDANCERCTRLBASE.dut ---- *)
TYPE _SCPAR_TM_WINDERDANCERCTRLBASE :
STRUCT
	XLINEVELDIAMCALC : BOOL;
	LRDANCERPOSRAMP : LREAL := 1;
	LRDANCERPOSCTRLGAIN : LREAL := 1;
	LRDANCERPOSCTRLRESETTIME : LREAL := 0;
	LRDANCERPOSCTRLLIMITPOS : LREAL := 1;
	LRDANCERPOSCTRLLIMITNEG : LREAL := -1;
	LRDANCERMAXPOSSCALED : LREAL := 0.95;
	LRDANCERMINPOSSCALED : LREAL := -0.95;
	XTEACHDANCERLIMITS : BOOL := FALSE;
	LRDANCERUPPERLIMIT : LREAL := 10000000;
	LRDANCERLOWERLIMIT : LREAL := 0;
	LRDANCERMATERIALLENGTH : LREAL := 0;
	LRDANCERINPOSWINDOWSCALED : LREAL := 0.2;
	RFILTTIMEACTDANCERPOSIN : REAL := 0.005;
	RFILTTIMEACTDANCERVELCOMP : REAL := 0;
	WWEBBREAKMODE : WORD := 1;
END_STRUCT
END_TYPE

(* ---- _SCPAR_TM_WINDERDANCERCTRLHIGH.dut ---- *)
TYPE _SCPAR_TM_WINDERDANCERCTRLHIGH :
STRUCT
	RFILTTIMEIDENTMINERTIASPD : REAL := 0.01;
	RFILTTIMEIDENTMINERTIATRQ : REAL := 0.005;
	LRIDENTMINERTIAMAXSPDSCALED : LREAL := 0.2;
	LRIDENTMINERTIAMAXTRQSCALED : LREAL := 0.2;
	EADAPTSPDCTRLGAINMODE : L_TT1P_AdaptSpdCtrlGainMode := 2;
	LRADAPTSPDCTRLLOWLIMIT : LREAL := 0;
	ALRSPDCTRLGAINADAPTX : ARRAY [1..9] OF LREAL := [0, 0.2, 0.4, 0.6, 0.8, 1, 1.2, 1.4, 1.6];
	ALRSPDCTRLGAINADAPTY : ARRAY [1..9] OF LREAL := [0.5, 0.6, 0.7, 0.8, 0.9, 1, 0.98, 0.95, 0.95];
	LRREDUCEDGAINWINDOW : LREAL;
	LRREDUCEDGAIN : LREAL;
	EDANCERCTRLSTOPMODE : L_TT1P_DancerCtrlStopMode;
	LRVEL : LREAL;
	LRACC : LREAL := 100;
	LRDEC : LREAL := 100;
	LRPOS_DIST : LREAL;
	LRIDENTDIAMVEL : LREAL := 10;
	LRIDENTDIAMACC : LREAL := 100;
	LRIDENTDIAMDEC : LREAL := 100;
	LRIDENTDIAMJERK : LREAL;
	WIDENTDIAMCALCCYCLES : WORD := 2;
	LRIDENTDIAMMAXDANCERPOS : LREAL := 0.5;
	LRIDENTDIAMSPDCTRLGAIN : LREAL := 0.5;
END_STRUCT
END_TYPE

(* ---- _SCPAR_TM_WINDERDANCERCTRLSTATE.dut ---- *)
TYPE _SCPAR_TM_WINDERDANCERCTRLSTATE :
STRUCT
	DWSELECTTENSCURVE : DWORD := 0;
	ALRTENSCURVE : ARRAY [1..65] OF LREAL;
	RFILTTIMEACCSPD : REAL := 0.005;
	LRACCCMPSDEADBANDTRQSCALED : LREAL := 0.1;
	LRACCCMPSGAINACC : LREAL := 1.05;
	LRACCCMPSGAINDEC : LREAL := 0.95;
	LRCONSTMINERTIA : LREAL := 9;
	LRMAXMINERTIA : LREAL := 50;
END_STRUCT
END_TYPE

(* ---- _SCPAR_TM_WINDERTENSIONCTRLBASE.dut ---- *)
TYPE _SCPAR_TM_WINDERTENSIONCTRLBASE :
STRUCT
	LRLINEVELOFFSETSCALED : LREAL := 0.1;
	LRTENSREF : LREAL := 2;
	LRTENSRAMP : LREAL := 1;
	RFILTTIMEWNDSPD : REAL := 0.01;
	RFILTTIMEACCSPD : REAL := 0.005;
	LRACCCMPSDEADBANDTRQSCALED : LREAL := 0.1;
	LRACCCMPSGAINACC : LREAL := 1.05;
	LRACCCMPSGAINDEC : LREAL := 0.95;
	LRCONSTMINERTIA : LREAL := 9;
	LRMAXMINERTIA : LREAL := 50;
	LRFRICCURVESTARTTRQ : LREAL := 0;
	LRFRICCURVEENDTRQ : LREAL := 0;
	RFILTTIMEFRICSETSPD : REAL := 0.01;
END_STRUCT
END_TYPE

(* ---- _SCPAR_TM_WINDERTENSIONCTRLHIGH.dut ---- *)
TYPE _SCPAR_TM_WINDERTENSIONCTRLHIGH :
STRUCT
	RFILTTIMEIDENTMINERTIASPD : REAL := 0.01;
	RFILTTIMEIDENTMINERTIATRQ : REAL := 0.005;
	LRIDENTMINERTIAMAXSPDSCALED : LREAL := 0.2;
	LRIDENTMINERTIAMAXTRQSCALED : LREAL := 0.2;
	EADAPTSPDCTRLGAINMODE : L_TT1P_AdaptSpdCtrlGainMode := 2;
	LRADAPTSPDCTRLLOWLIMIT : LREAL := 0;
	ALRSPDCTRLGAINADAPTX : ARRAY [1..9] OF LREAL := [0, 0.2, 0.4, 0.6, 0.8, 1, 1.2, 1.4, 1.6];
	ALRSPDCTRLGAINADAPTY : ARRAY [1..9] OF LREAL := [0.5, 0.6, 0.7, 0.8, 0.9, 1, 0.98, 0.95, 0.95];
	LRREDUCEDGAINWINDOW : LREAL;
	LRREDUCEDGAIN : LREAL;
	ETENSCTRLSTOPMODE : L_TT1P_TensionCtrlStopMode;
	LRVEL : LREAL;
	LRACC : LREAL := 100;
	LRDEC : LREAL := 100;
	LRPOS_DIST : LREAL;
END_STRUCT
END_TYPE

(* ---- _SCPAR_TM_WINDERTENSIONCTRLSTATE.dut ---- *)
TYPE _SCPAR_TM_WINDERTENSIONCTRLSTATE :
STRUCT
	DWSELECTTENSCURVE : DWORD := 0;
	ALRTENSCURVE : ARRAY [1..65] OF LREAL;
	LRTENSCTRLGAIN : LREAL := 0;
	LRTENSCTRLRESETTIME : LREAL := 0;
	LRTENSCTRLLIMITPOS : LREAL := L_UMTP_Math.gC_POSITIVE_LIMIT_32BIT;
	LRTENSCTRLLIMITNEG : LREAL := L_UMTP_Math.gC_NEGATIVE_LIMIT_32BIT;
	LRIDENTFRICMAXSPDSCALED : LREAL := 0.9;
	LRIDENTFRICACCDEC : LREAL := 1;
	RFILTTIMEIDENTFRICSPD : REAL := 0.0;
	RFILTTIMEIDENTFRICTRQ : REAL := 0.05;
	DWSELECTFRICCURVE : DWORD := 1;
	RFILTTIMEACTTENSIN : REAL := 0.005;
	LRACTTENSINGAIN : LREAL := 1;
	LRACTTENSINOFFSET : LREAL := 0;
END_STRUCT
END_TYPE

(* ---- _SCSF_TM_BASICMOTIONBASE.dut ---- *)
TYPE _SCSF_TM_BASICMOTIONBASE :
STRUCT
END_STRUCT
END_TYPE

(* ---- _SCSF_TM_BASICMOTIONHIGH.dut ---- *)
TYPE _SCSF_TM_BASICMOTIONHIGH :
STRUCT
END_STRUCT
END_TYPE

(* ---- _SCSF_TM_BASICMOTIONSTATE.dut ---- *)
TYPE _SCSF_TM_BASICMOTIONSTATE :
STRUCT
END_STRUCT
END_TYPE

(* ---- _SCSF_TM_CROSSCUTTERBASE.dut ---- *)
TYPE _SCSF_TM_CROSSCUTTERBASE :
STRUCT
	IP01_ECUTTINGMODE : L_TT1P_CuttingModeState;
	IP02_LRSCALINGMASTER : LREAL;
	IP03_LRSETOFFSETMASTER : LREAL;
	MP00_LWCHECKSUMENDOFPROFILE : LWORD;
	MP01_LRSETMASTERPOS : LREAL;
	MP02_LRCAMPROFILERPOSOUT : LREAL;
	MP03_LRSETSLAVEPOSOUT : LREAL;
	MP04_CAMPOINTSTART : ARRAY [0..3] OF L_MC2P_CamDataXYVA;
	MP05_CAMPOINTCONTINUOUS : ARRAY [0..5] OF L_MC2P_CamDataXYVA;
	MP06_CAMPOINTSTOP : ARRAY [0..3] OF L_MC2P_CamDataXYVA;
	MP07_INUMOFPOINTSINCAM : INT;
	MP08_BYSELECTCAM : BYTE;
	MP09_ECUTTINGPROCESSSTATE : L_TT1P_States;
	MP10_LRYSTART : LREAL;
	MP11_LRYPARK : LREAL;
	MP12_LRYEND : LREAL;
	MP13_LRXSTART : LREAL;
	MP14_LRXENDSYNCPOS : LREAL;
	MP15_LRXSTARTPARKPOS : LREAL;
	MP16_LRXENDPARKPOS : LREAL;
	MP17_LRXSTARTSYNCPOS : LREAL;
	MP18_LRXEND : LREAL;
	MP19_XXABSOLUTE : BOOL;
	MP20_XSLAVEABSOLUTE : BOOL;
	MP21_XENDOFPROFILE : BOOL;
	MP22_XENDOFXCYCLE : BOOL;
	MP23_XENABLEPOSITIONFOLLOWER : BOOL;
	MP24_LRSETOVERSPEEDSCALED : LREAL;
	AP01_XENDOFPROFILEWINDOWSIZE : BOOL;
	AP01_LRENDOFPROFILEWINDOWSIZE : LREAL := 0;
	AP02_XOVERSPEEDUPPERLIMIT : BOOL;
	AP02_LROVERSPEEDUPPERLIMIT : LREAL := 2;
END_STRUCT
END_TYPE

(* ---- _SCSF_TM_CROSSCUTTERHIGH.dut ---- *)
TYPE _SCSF_TM_CROSSCUTTERHIGH :
STRUCT
END_STRUCT
END_TYPE

(* ---- _SCSF_TM_CROSSCUTTERSTATE.dut ---- *)
TYPE _SCSF_TM_CROSSCUTTERSTATE :
STRUCT
	IP04_LRMINERTIA : LREAL;
	IP05_XMARKRECEIVE : BOOL;
	IP06_LRACTMARKPOSIN : LREAL;
	IP07_LRMAXCORRPOS : LREAL;
	IP08_LRMAXCORRNEG : LREAL;
	IP09_XMARKCORRECTION : BOOL;
	MP25_XENABLETORQUEFOLLOWER : BOOL;
	MP26_LRPRECTRLACCOUT : LREAL;
	MP27_LRGEARBOXFACTOR : LREAL;
	MP28_LRAXISTORQUE : LREAL;
	MP30_LRSETVELOCITYREGISTER : LREAL;
	MP31_LRINTEGRATORREGPOS : LREAL;
	MP32_LRCORRREGPOS : LREAL;
	MP33_LRMARKSENSORPOS : LREAL;
	MP34_XMARKRECEIVEUNLIMITED : BOOL;
	MP35_LRACTMARKERRORUNLIMITED : LREAL;
	MP36_LRUPPERCORRPOS : LREAL;
	MP37_LRLOWERCORRPOS : LREAL;
	MP38_LRMARKDIST : LREAL;
	OP02_LRSETMOTORPRECTRLTRQOUT : LREAL;
	OP03_LRREGMARKPOS : LREAL;
	OP04_XMARKRECEIVED : BOOL;
	OP05_LRACTMARKERROR : LREAL;
	OP06_LRSETREGPOSOUT : LREAL;
	AP03_XTPAXISDELAYCYCLE : BOOL;
	AP03_LRTPAXISDELAYCYCLE : LREAL;
	AP04_XTPAXISCOMPFACTOR : BOOL;
	AP04_LRTPAXISCOMPFACTOR : LREAL;
	AP05_XUPPERCORRPOS : BOOL;
	AP05_LRUPPERCORRPOS : LREAL;
	AP06_XLOWERCORRPOS : BOOL;
	AP06_LRLOWERCORRPOS : LREAL;
END_STRUCT
END_TYPE

(* ---- _SCSF_TM_ELECTRICALSHAFTPOSBASE.dut ---- *)
TYPE _SCSF_TM_ELECTRICALSHAFTPOSBASE :
STRUCT
	IP01_LRSETOFFSETSLAVE : LREAL;
	AP01_XLOADGEARBOXPOSOUT : BOOL;
	AP01_LRLOADGEARBOXPOSOUT : LREAL;
	MP01_LRSETMASTERPOS : LREAL;
	MP02_LRSETSLAVEPOS : LREAL;
	MP03_LRSETGEARBOXPOSOUT : LREAL;
	OP01_LROFFSET : LREAL;
END_STRUCT
END_TYPE

(* ---- _SCSF_TM_ELECTRICALSHAFTPOSHIGH.dut ---- *)
TYPE _SCSF_TM_ELECTRICALSHAFTPOSHIGH :
STRUCT
	IP02_LRSETOFFSETMASTER : LREAL;
	OP04_LROFFSETMASTER : LREAL;
END_STRUCT
END_TYPE

(* ---- _SCSF_TM_ELECTRICALSHAFTPOSSTATE.dut ---- *)
TYPE _SCSF_TM_ELECTRICALSHAFTPOSSTATE :
STRUCT
	AP02_XLOADTRIMOFFSET : BOOL;
	AP02_LRLOADTRIMOFFSET : LREAL;
	MP04_LRSETCLUTCHPOS : LREAL;
	OP02_LROFFSETTRIM : LREAL;
	OP03_LROFFSETTOTAL : LREAL;
END_STRUCT
END_TYPE

(* ---- _SCSF_TM_ELECTRICALSHAFTVELBASE.dut ---- *)
TYPE _SCSF_TM_ELECTRICALSHAFTVELBASE :
STRUCT
	AP01_XCOUPLINGX : BOOL;
	AP01_LRCOUPLINGX : LREAL := 1.0;
	AP02_XCOUPLINGY : BOOL;
	AP02_LRCOUPLINGY : LREAL := 1.0;
	IP01_LRSETOFFSETSLAVE : LREAL;
	MP01_LRSETMASTERVEL : LREAL;
	MP02_LRSETCLUTCHVEL : LREAL;
	MP03_LRSETSLAVEVEL : LREAL;
	MP04_LRSETGEARBOXOUTVEL : LREAL;
	OP01_LROFFSET : LREAL;
END_STRUCT
END_TYPE

(* ---- _SCSF_TM_ELECTRICALSHAFTVELHIGH.dut ---- *)
TYPE _SCSF_TM_ELECTRICALSHAFTVELHIGH :
STRUCT
END_STRUCT
END_TYPE

(* ---- _SCSF_TM_ELECTRICALSHAFTVELSTATE.dut ---- *)
TYPE _SCSF_TM_ELECTRICALSHAFTVELSTATE :
STRUCT
	OP02_LROFFSETTRIM : LREAL;
	OP03_LROFFSETTOTAL : LREAL;
END_STRUCT
END_TYPE

(* ---- _SCSF_TM_FLEXCAMBASE.dut ---- *)
TYPE _SCSF_TM_FLEXCAMBASE :
STRUCT
	IP01_LRSETSCALINGMASTER : LREAL;
	IP02_ESCALINGMODEMASTER : L_TT1P_ScalingMode;
	IP03_LRSETOFFSETMASTER : LREAL;
	IP04_LRSETOFFSETSLAVE : LREAL;
	IP05_EOFFSETMODESLAVE : L_TT1P_OffsetModeSlave;
	IP06_LRSETSCALINGSLAVE : LREAL;
	IP07_ESCALINGMODESLAVE : L_TT1P_ScalingMode;
	IP08_CAMTABLE1 : MC_CAM_REF;
	MP01_LRSETMASTERPOS : LREAL;
	MP02_LRSETSLAVEPOS : LREAL;
	MP03_LRCONVERTMASTERTOXPOS : LREAL;
	MP04_LRCAMPROFILERPOSOUT : LREAL;
	MP05_LRSETYPOS : LREAL;
	MP06_LRCONVERTYTOSLAVEPOS : LREAL;
	MP07_XENDOFPROFPOSITIVE : BOOL;
	MP08_XENDOFPROFNEGATIVE : BOOL;
	OP01_LRSETXPOSOUT : LREAL;
	OP02_LESETYPOSOUT : LREAL;
	MP00_LWENDOFPROFILECHECKSUM : LWORD;
END_STRUCT
END_TYPE

(* ---- _SCSF_TM_FLEXCAMHIGH.dut ---- *)
TYPE _SCSF_TM_FLEXCAMHIGH :
STRUCT
END_STRUCT
END_TYPE

(* ---- _SCSF_TM_FLEXCAMSTATE.dut ---- *)
TYPE _SCSF_TM_FLEXCAMSTATE :
STRUCT
	IP09_CAMTABLE2 : MC_CAM_REF;
	IP10_CAMTABLE3 : MC_CAM_REF;
	IP11_CAMTABLE4 : MC_CAM_REF;
END_STRUCT
END_TYPE

(* ---- _SCSF_TM_FLYINGSAWBASE.dut ---- *)
TYPE _SCSF_TM_FLYINGSAWBASE :
STRUCT
	IP01_XEXECUTENEXTCUT : BOOL;
	IP02_LRCUTTINGLENGTH : LREAL;
	IP03_LRLOWERLIMIT : LREAL;
	IP04_LRUPPERLIMIT : LREAL;
	AP01_XLOADTOTALCUTTINGLENGTH : BOOL;
	AP01_LRLOADTOTALCUTTINGLENGTH : LREAL;
	AP02_XLOADTARGETPOS : BOOL;
	AP02_LRLOADTARGETPOS : LREAL;
	MP01_LRSETMASTERPOS : LREAL;
	MP02_LRSETSLAVEPOS : LREAL;
	MP03_LRTOTALCUTTINGLENGTH : LREAL;
	MP04_XPOSSYNCHRONISED : BOOL;
	OP01_LRMATERIALCOUNTER : LREAL;
	OP02_LRTARGETPOS : LREAL;
END_STRUCT
END_TYPE

(* ---- _SCSF_TM_FLYINGSAWHIGH.dut ---- *)
TYPE _SCSF_TM_FLYINGSAWHIGH :
STRUCT
END_STRUCT
END_TYPE

(* ---- _SCSF_TM_FLYINGSAWSTATE.dut ---- *)
TYPE _SCSF_TM_FLYINGSAWSTATE :
STRUCT
	IP05_EMODEFLYINGSAW : L_TT1P_eModesFlyingSaw;
	AP03_XRANGEOFTOLERANCE : BOOL;
	AP03_LRRANGEOFTOLERANCE : LREAL;
	AP04_XMARKDETECTERRCOMP : BOOL;
	AP04_LRMARKDETECTERRCOMP : LREAL;
	MP05_WMARKININDEX : WORD;
	MP06_WMARKOUTINDEX : WORD;
	MP07_ALRMARKPOSITIONARRAY : ARRAY [0..15] OF LREAL;
	MP08_ALRTIMESTAMPARRAY : ARRAY [0..15] OF LREAL;
	MP09_XMARKSTACKEMPTY : BOOL;
	MP10_XMARKSTACKFULL : BOOL;
	MP11_MARKPOS : LREAL;
END_STRUCT
END_TYPE

(* ---- _SCSF_TM_MOTIONCONTROL.dut ---- *)
TYPE _SCSF_TM_MOTIONCONTROL :
STRUCT
	MP00_LWTCHECKSUM : LWORD;
END_STRUCT
END_TYPE

(* ---- _SCSF_TM_PICKANDPLACEBASE.dut ---- *)
TYPE _SCSF_TM_PICKANDPLACEBASE :
STRUCT
	MP00_LWTCHECKSUM : LWORD;
	MP01_LRSETA1POS : LREAL;
	MP02_LRSETA2POS : LREAL;
	MP03_LRSETA3POS : LREAL;
	MP04_LRSETA4POS : LREAL;
	MP05_LRSTARTXPOS : LREAL;
	MP06_LRSTARTYPOS : LREAL;
	MP07_LRSTARTZPOS : LREAL;
	MP08_LRSTARTAUX1POS : LREAL;
	MP09_LRSETXPOS : LREAL;
	MP10_LRSETYPOS : LREAL;
	MP11_LRSETZPOS : LREAL;
	MP12_LRSETAUX1POS : LREAL;
	MP13_BYINTERMEDIANTEPOINT : BYTE;
	MP15_DISEGMENTNO : DINT;
	MP20_PAMOVELINEARABSOLUTE : POINTER TO ARRAY [1..10] OF MC_MoveLinearAbsolute;
END_STRUCT
END_TYPE

(* ---- _SCSF_TM_PICKANDPLACEHIGH.dut ---- *)
TYPE _SCSF_TM_PICKANDPLACEHIGH :
STRUCT
	MP21_PAMOVELINEARABSOLUTE : POINTER TO ARRAY [1..10] OF L_MC4P_MoveLinearAbsolute_Internal;
	MP22_PAMOVELINEARABSOLUTE : POINTER TO ARRAY [1..10] OF L_MC4P_MoveLinearAbsolute_Internal;
	MP23_PAMOVELINEARABSOLUTE : POINTER TO ARRAY [1..10] OF L_MC4P_MoveLinearAbsolute_Internal;
	MP25_IMOVEPPNO : INT;
	MP26_IMOVELINNO : INT;
END_STRUCT
END_TYPE

(* ---- _SCSF_TM_PICKANDPLACESTATE.dut ---- *)
TYPE _SCSF_TM_PICKANDPLACESTATE :
STRUCT
	MP14_ALRINTERMEDIANTEPOINT : ARRAY [1..12] OF LREAL;
END_STRUCT
END_TYPE

(* ---- _SCSF_TM_REGISTERCONTROLBASE.dut ---- *)
TYPE _SCSF_TM_REGISTERCONTROLBASE :
STRUCT
	IP01_LRSETMASTERPOS : LREAL;
	IP02_XLOADREGISTERPOS : BOOL;
	IP03_LRMARKDIST : LREAL;
	IP04_XMARKRECEIVE : BOOL;
	IP05_LRACTMARKPOSIN : LREAL;
	IP06_LRMAXCORRPOS : LREAL;
	IP07_LRMAXCORRNEG : LREAL;
	IP08_LRUPPERCORRPOS : LREAL;
	IP09_LRLOWERCORRPOS : LREAL;
	IP10_XMARKCORR : BOOL;
	IP11_LRSLAVEAXISCYCLELENGTH : LREAL;
	IP12_ETRIMMODE : L_TT1P_TrimMode;
	IP13_LRSETOFFSETMASTER : LREAL;
	IP14_DWDENOMINATOR : DWORD;
	IP15_DWNUMERATOR : DWORD;
	IP16_LRMASTERAXISCYCLELENGTH : LREAL;
	IP17_LRSETOFFSETSLAVE : LREAL;
	MP01_LRSETVELOCITYREGISTER : LREAL;
	MP02_LRINTEGRATORREGPOS : LREAL;
	MP03_LRCORRREGPOS : LREAL;
	MP04_LRMARKSENSORPOS : LREAL;
	MP05_XMARKRECEIVEUNLIMITED : BOOL;
	MP06_LRACTMARKERRORUNLIMITED : LREAL;
	MP07_LRSETGEARBOXPOSIN : LREAL;
	MP08_LRSETGEARBOXPOSOUT : LREAL;
	MP09_LRSETCLUTCHPOSIN : LREAL;
	OP01_LRREGPOSOUT : LREAL;
	OP02_LRREGMARKPOS : LREAL;
	OP03_XMARKRECEIVED : BOOL;
	OP04_LRACTMARKERROR : LREAL;
	AP03_XTPAXISDELAYCYCLE : BOOL;
	AP03_LRTPAXISDELAYCYCLE : LREAL;
	AP04_XTPAXISCOMPFACTOR : BOOL;
	AP04_LRTPAXISCOMPFACTOR : LREAL;
END_STRUCT
END_TYPE

(* ---- _SCSF_TM_REGISTERCONTROLHIGH.dut ---- *)
TYPE _SCSF_TM_REGISTERCONTROLHIGH :
STRUCT
END_STRUCT
END_TYPE

(* ---- _SCSF_TM_REGISTERCONTROLSTATE.dut ---- *)
TYPE _SCSF_TM_REGISTERCONTROLSTATE :
STRUCT
	IP18_XGEARFACTORCORR : BOOL;
	IP19_LRMARKWINDOWSIZE : LREAL;
	IP20_DWMISSEDMARKS : DWORD;
	IP21_XTEACHMARKWINDOW : BOOL;
	MP10_XMARKWINDOWCOMPOUT : BOOL;
	MP11_LRMARKSTACKLENGTH : LREAL;
	MP12_LRMARKSTACKERRORTOTAL : LREAL;
	MP13_XMARKRECEIVEDLIMITED : BOOL;
	MP14_LRACTMARKERRORLIMITED : LREAL;
END_STRUCT
END_TYPE

(* ---- _SCSF_TM_SMARTTRACKBASE.dut ---- *)
TYPE _SCSF_TM_SMARTTRACKBASE :
STRUCT
END_STRUCT
END_TYPE

(* ---- _SCSF_TM_SMARTTRACKHIGH.dut ---- *)
TYPE _SCSF_TM_SMARTTRACKHIGH :
STRUCT
END_STRUCT
END_TYPE

(* ---- _SCSF_TM_SMARTTRACKSTATE.dut ---- *)
TYPE _SCSF_TM_SMARTTRACKSTATE :
STRUCT
	MP01_ALRPRODUCTPOSITION : ARRAY [1..10] OF LREAL;
END_STRUCT
END_TYPE

(* ---- _SCSF_TM_STACKERCRANEAXISCONTROLBASE.dut ---- *)
TYPE _SCSF_TM_STACKERCRANEAXISCONTROLBASE :
STRUCT
	MP01_LROSCCOMPLOADSCALED : LREAL;
	MP02_LROSCCOMPPOSSCALED : LREAL;
	MP03_LROSCCOMPAMPRATIO : LREAL;
	MP04_LROSCCOMPEIGENFREQ : LREAL;
	MP05_XOSCCOMPBUSY : BOOL;
	MP06_XOSCCOMPINEQOUT : BOOL;
	MP07_XOSCCOMPACTIVE : BOOL;
	MP08_LROSCCOMPSETPOSOUT : LREAL;
	MP09_LROSCCOMPSETVELOUT : LREAL;
	MP10_LROSCCOMPSETACCOUT : LREAL;
	MP11_LROSCCOMPSETTORQUEOUT : LREAL;
	MP12_XBRAKEGRINDINBUSY : BOOL;
	MP13_XBRAKEGRINDINACTIVE : BOOL;
	MP14_XBRAKEGRINDINDONE : BOOL;
	MP15_XBRAKETESTBUSY : BOOL;
	MP16_XBRAKETESTACTIVE : BOOL;
	MP17_XBRAKETESTDONE : BOOL;
	MP18_LRBRAKETESTIDENTTORQUE : LREAL;
	MP19_LRBRAKETESTACTPOSTHRESHOLD : LREAL;
	MP20_LRBRAKETESTACTMOTORTORQUE : LREAL;
	MP21_XIDENTCONSTTORQUEVALID : BOOL;
	MP22_LRIDENTCONSTTORQUE : LREAL;
	MP23_LRFILTACTTORQUE : LREAL;
END_STRUCT
END_TYPE

(* ---- _SCSF_TM_STACKERCRANEHEADCONTROLBASE.dut ---- *)
TYPE _SCSF_TM_STACKERCRANEHEADCONTROLBASE :
STRUCT
	MP01_XCOMMUNICATIONVALID : BOOL;
	MP02_XLOCKCOMCHANNEL : BOOL;
	MP10_XPROFILEDATAXVALID : BOOL;
	MP11_SCPROFILEDATAX : L_TT1P_ProfileGeneratorData;
	MP12_SCBUFFPROFILEDATAX : L_TT1P_ProfileGeneratorData;
	MP13_XPROFILEDATAYVALID : BOOL;
	MP14_SCPROFILEDATAY : L_TT1P_ProfileGeneratorData;
	MP15_SCBUFFPROFILEDATAY : L_TT1P_ProfileGeneratorData;
END_STRUCT
END_TYPE

(* ---- _SCSF_TM_TABLEPOSITIONINGBASE.dut ---- *)
TYPE _SCSF_TM_TABLEPOSITIONINGBASE :
STRUCT
END_STRUCT
END_TYPE

(* ---- _SCSF_TM_TABLEPOSITIONINGHIGH.dut ---- *)
TYPE _SCSF_TM_TABLEPOSITIONINGHIGH :
STRUCT
END_STRUCT
END_TYPE

(* ---- _SCSF_TM_TABLEPOSITIONINGSTATE.dut ---- *)
TYPE _SCSF_TM_TABLEPOSITIONINGSTATE :
STRUCT
END_STRUCT
END_TYPE

(* ---- _SCSF_TM_WINDER.dut ---- *)
TYPE _SCSF_TM_WINDER :
STRUCT
	AP10_XSETTRQOFFSET : BOOL;
	AP10_LRSETTRQOFFSET : LREAL;
	AP09_XSETVELOFFSET : BOOL;
	AP09_LRSETVELOFFSET : LREAL;
	MP15_LRWNDVELREF : LREAL;
	MP16_LRWNDSPEEDREF : LREAL;
	MP20_LIREVCOUNTER : LINT;
	MP21_LRREVCOUNTERRESIDUAL : LREAL;
	MP22_LRAXISSPEED : LREAL;
END_STRUCT
END_TYPE

(* ---- _SCSF_TM_WINDERDANCERCTRLBASE.dut ---- *)
TYPE _SCSF_TM_WINDERDANCERCTRLBASE :
STRUCT
	IP01_LRSETLINEVEL : LREAL;
	IP02_LRSETLINEVELDIAMCALC : LREAL;
	IP03_XLINEVELDIAMCALC : BOOL;
	IP04_LRDANCERMATERIALLENGTH : LREAL;
	IP05_LRSETDIAM : LREAL;
	IP06_XLOADDIAM : BOOL;
	IP07_XWINDINGDIRECTION : BOOL;
	IP08_XMATERIALFEEDING : BOOL;
	IP09_LRACTDANCERPOSIN : LREAL;
	IP10_LRSETDANCERPOSSCALED : LREAL;
	IP11_LRLINEVELREF : LREAL;
	IP12_LRSETTENS : LREAL;
	AP01_XSETSPEEDPOINT : BOOL;
	AP01_LRSETSPEEDPOINT : LREAL;
	AP03_XSETDANCERCTRLOUTGAIN : BOOL;
	AP03_LRSETDANCERCTRLOUTGAIN : LREAL;
	AP04_XSETDANCERCTRLOUTRESETTIME : BOOL;
	AP04_LRSETDANCERCTRLOUTRESETTIME : LREAL;
	AP05_XSETDANCERCTRLOUTRATETIME : BOOL;
	AP05_LRSETDANCERCTRLOUTRATETIME : LREAL;
	MP01_LRDANCERPOSSCALED0TO1 : LREAL;
	MP02_LRDANCERCOMPVELOUT : LREAL;
	MP03_LRFILTDANCERCOMPVELOUT : LREAL;
	MP04_LRFILTACTDANCERPOSSCALED : LREAL;
	MP05_LRSETRAMPDANCERPOS : LREAL;
	MP06_LRDANCERCTRLPOSOUT : LREAL;
	MP06_1_LRPDANCERCTRLOUT : LREAL;
	MP06_2_LRIDANCERCTRLOUT : LREAL;
	MP06_3_LRDDANCERCTRLOUT : LREAL;
	MP07_LRDANCERCTRLLINEVELOUT : LREAL;
	MP08_LRSETSPEEDPOINT : LREAL;
	MP11_LRDANCERCTRLOUTGAIN : LREAL;
	MP12_LRDANCERCTRLOUTRESETTIME : LREAL;
	MP13_LRDANCERCTRLOUTRATETIME : LREAL;
	OP01_LRACTDANCERPOSSCALED : LREAL;
	OP02_LRSETDIAMOUT : LREAL;
	OP03_LRAXISSPEED : LREAL;
	OP04_LRSETTENSCURVEOUT : LREAL;
END_STRUCT
END_TYPE

(* ---- _SCSF_TM_WINDERDANCERCTRLHIGH.dut ---- *)
TYPE _SCSF_TM_WINDERDANCERCTRLHIGH :
STRUCT
END_STRUCT
END_TYPE

(* ---- _SCSF_TM_WINDERDANCERCTRLSTATE.dut ---- *)
TYPE _SCSF_TM_WINDERDANCERCTRLSTATE :
STRUCT
	AP02_XSETTRQPOINT : BOOL;
	AP02_LRSETTRQPOINT : LREAL;
	MP09_LRAXISTORQUE : LREAL;
	MP10_LRSETTRQPOINT : LREAL;
END_STRUCT
END_TYPE

(* ---- _SCSF_TM_WINDERTENSIONCTRLBASE.dut ---- *)
TYPE _SCSF_TM_WINDERTENSIONCTRLBASE :
STRUCT
	IP01_LRSETLINEVEL : LREAL;
	IP02_LRSETDIAM : LREAL;
	IP03_XLOADDIAM : BOOL;
	IP04_LRLINEVELOFFSETSCALED : LREAL;
	IP05_LRLINEVELREF : LREAL;
	IP06_XMATERIALFEEDING : BOOL;
	IP07_LRSETTENSION : LREAL;
	IP08_XWINDINGDIRECTION : BOOL;
	AP01_XSETACCCOMPTRQ : BOOL;
	AP01_LRSETACCCOMPTRQ : LREAL;
	AP02_XSETTRQPOINT : BOOL;
	AP02_LRSETTRQPOINT : LREAL;
	AP03_XSETUPPERSPEEDLIMIT : BOOL;
	AP03_LRSETUPPERSPEEDLIMIT : LREAL;
	AP04_XSETLOWERSPEEDLIMIT : BOOL;
	AP04_LRSETLOWERSPEEDLIMIT : LREAL;
	MP01_LRTENSCURVEOUT : LREAL;
	MP02_LRSETTENSPOINT : LREAL;
	MP03_LRSETTENSTRQ : LREAL;
	MP04_LRSETACCCOMPTRQ : LREAL;
	MP05_LRSETFRICCOMPTRQ : LREAL;
	MP06_LRSETTRQPOINT : LREAL;
	MP07_LRSETUPPERSPEEDLIMIT : LREAL;
	MP08_LRSETLOWERSPEEDLIMIT : LREAL;
	MP09_LRAXISUPPERSPEEDLIMIT : LREAL;
	MP10_LRAXISLOWERSPEEDLIMIT : LREAL;
	MP11_LRAXISVEL : LREAL;
	MP12_LRAXISTORQUE : LREAL;
	OP01_LRSETDIAMOUT : LREAL;
END_STRUCT
END_TYPE

(* ---- _SCSF_TM_WINDERTENSIONCTRLHIGH.dut ---- *)
TYPE _SCSF_TM_WINDERTENSIONCTRLHIGH :
STRUCT
END_STRUCT
END_TYPE

(* ---- _SCSF_TM_WINDERTENSIONCTRLSTATE.dut ---- *)
TYPE _SCSF_TM_WINDERTENSIONCTRLSTATE :
STRUCT
	IP09_LRACTTENSIN : LREAL;
	MP13_LRFILTACTTENSIN : LREAL;
	MP14_LRTENSCTRLOUT : LREAL;
	MP15_LRPTENSCTRLOUT : LREAL;
	MP16_LRITENSCTRLOUT : LREAL;
	MP17_LRDTENSCTRLOUT : LREAL;
	MP15_LRTENSCTRLOUTGAIN : LREAL;
	MP16_LRTENSCTRLOUTRESETTIME : LREAL;
	MP17_LRTENSCTRLOUTRATETIME : LREAL;
	MP18_LRSETTENSCTRLVALUE : LREAL;
	MP19_LRACTTENSCTRLVALUE : LREAL;
	AP05_XSETTENSIONCTRLOUTGAIN : BOOL;
	AP05_LRSETTENSIONCTRLOUTGAIN : LREAL;
	AP06_XSETTENSIONCTRLOUTRESETTIME : BOOL;
	AP06_LRSETTENSIONCTRLOUTRESETTIME : LREAL;
	AP07_XSETTENSIONCTRLOUTRATETIME : BOOL;
	AP07_LRSETTENSIONCTRLOUTRATETIME : LREAL;
	AP08_XSETFRICCOMPREELSPEED : BOOL;
	AP08_LRSETFRICCOMPREELSPEED : LREAL;
END_STRUCT
END_TYPE

(* ---- L_MB1P_AXISPROFILE.dut ---- *)
TYPE L_MB1P_AXISPROFILE :
STRUCT
	LRPOS : LREAL;
	LRVEL : LREAL;
	LRACC : LREAL;
END_STRUCT
END_TYPE

(* ---- L_MB1P_CAMSEQUENCEMODE.dut ---- *)
TYPE L_MB1P_CAMSEQUENCEMODE :
(
	CYCLICCAM1 := 0,
	CYCLICCAM3 := 1,
	CAM1_CYCLICCAM3_CAM1 := 2,
	CAM1_CAM2_CYCLICCAM3_CAM4_CAM1 := 3
);
END_TYPE

(* ---- L_MB1P_CAMTABLE.dut ---- *)
TYPE L_MB1P_CAMTABLE :
(
	NOCAMTABLE := 0,
	CAMTABLE1 := 1,
	CAMTABLE2 := 2,
	CAMTABLE3 := 3,
	CAMTABLE4 := 4
);
END_TYPE

(* ---- L_MB1P_CHANNELDATA.dut ---- *)
TYPE L_MB1P_CHANNELDATA :
STRUCT
	XMASTER : BOOL;
	XSLAVE : BOOL;
	DWSTATUSWORD : DWORD;
	DWCONTROLWORD : DWORD;
	ETMSTATE : WORD;
	ALRDATA : ARRAY [1..20] OF LREAL;
	AIDATA : ARRAY [1..5] OF INT;
	ADWDATA : ARRAY [1..5] OF DWORD;
	XPOINTERTOAXISVALID : BOOL;
	PAXIS : POINTER TO AXIS_REF;
END_STRUCT
END_TYPE

(* ---- L_MB1P_CHANNELELEMENT.dut ---- *)
TYPE L_MB1P_CHANNELELEMENT :
STRUCT
	ITFCOMID : ITF_DataBus;
	XVALID : BOOL;
	DWMASK : DWORD;
	IELEMENTNO : INT := 1;
	ILEFT : INT := 1;
	IRIGHT : INT := 1;
	PLEFT : POINTER TO L_MB1P_ChannelElement;
	PRIGHT : POINTER TO L_MB1P_ChannelElement;
	PDATA : POINTER TO L_MB1P_ChannelData;
	PHEAD : POINTER TO L_MB1P_ChannelHeadData;
END_STRUCT
END_TYPE

(* ---- L_MB1P_CHANNELHEADDATA.dut ---- *)
TYPE L_MB1P_CHANNELHEADDATA :
STRUCT
	ICALLNUM : INT;
END_STRUCT
END_TYPE

(* ---- L_MB1P_CHARACTERISTICS.dut ---- *)
TYPE L_MB1P_CHARACTERISTICS :
STRUCT
	ELAWOFMOTIONCHAR : L_MB1P_LawOfMotionChar;
	LRX : LREAL;
	LRY : LREAL;
	LRA1 : LREAL;
	LRA2 : LREAL;
	LRA3 : LREAL;
	LRA4 : LREAL;
	LRA5 : LREAL;
END_STRUCT
END_TYPE

(* ---- L_MB1P_CLUTCHDIRECTION.dut ---- *)
TYPE L_MB1P_CLUTCHDIRECTION :
(
	MCNEGATIVEDIRECTION := -1,
	MCCURRENTDIRECTION := 0,
	MCPOSITIVEDIRECTION := 1
);
END_TYPE

(* ---- L_MB1P_CLUTCHMODE.dut ---- *)
TYPE L_MB1P_CLUTCHMODE :
(
	ABSOLUTE := 0,
	RELATIVE := 1,
	RAMP_POS := 2,
	RAMP_TIME := 3,
	RAMP_SLAVE_DIST := 4,
	ABSOLUTE_IN_TARGET := 5,
	RAMP_VELACC := 6,
	RAMP_RELATIVE := 7
);
END_TYPE

(* ---- L_MB1P_DATAPOINTSXY.dut ---- *)
TYPE L_MB1P_DATAPOINTSXY :
STRUCT
	LRX : LREAL;
	LRY : LREAL;
END_STRUCT
END_TYPE

(* ---- L_MB1P_DIRECTION.dut ---- *)
TYPE L_MB1P_DIRECTION :
(
	BOTH := 0,
	DIRECTIONMASTER := 1
);
END_TYPE

(* ---- L_MB1P_GCODELINE.dut ---- *)
TYPE L_MB1P_GCODELINE :
STRUCT
	G1 : BOOL;
	X : LREAL;
	Y : LREAL;
	Z : LREAL;
	C : LREAL;
	VELOCITY : LREAL;
	ACCELERATION : LREAL;
	DECELERATION : LREAL;
	G50 : BOOL;
	G51 : BOOL;
	D : LREAL;
	G70 : BOOL;
	G71 : BOOL;
	M1 : BOOL;
END_STRUCT
END_TYPE

(* ---- L_MB1P_INTPROFILEDATA.dut ---- *)
TYPE L_MB1P_INTPROFILEDATA :
STRUCT
	PHASE1 : L_MB1P_ProfilePhaseData;
	PHASE2 : L_MB1P_ProfilePhaseData;
	PHASE3 : L_MB1P_ProfilePhaseData;
	PHASE5 : L_MB1P_ProfilePhaseData;
	PHASE6 : L_MB1P_ProfilePhaseData;
	PHASE7 : L_MB1P_ProfilePhaseData;
END_STRUCT
END_TYPE

(* ---- L_MB1P_INTPROFILEDATAACC.dut ---- *)
TYPE L_MB1P_INTPROFILEDATAACC :
STRUCT
	PHASE1 : L_MB1P_ProfilePhaseData;
	PHASE2 : L_MB1P_ProfilePhaseData;
	PHASE3 : L_MB1P_ProfilePhaseData;
END_STRUCT
END_TYPE

(* ---- L_MB1P_LAWOFMOTIONCHAR.dut ---- *)
TYPE L_MB1P_LAWOFMOTIONCHAR :
(
	BB_POLY5 := 0,
	GG_MODSIN,
	GU_HARMKOMB,
	RR_BESCHLTRAPEZ,
	RR_GENSIN,
	RR_GERADE,
	RR_MODBESCHLTRAPEZ,
	RR_MODSIN,
	RR_POLY5,
	RR_QUADPARABEL,
	RR_SINUS,
	RU_MODBESCHLTRAPEZ,
	UG_HARMKOMB,
	UR_MODBESCHLTRAPEZ,
	UU_SINGERADEKOMB
);
END_TYPE

(* ---- L_MB1P_PROFILEDATA.dut ---- *)
TYPE L_MB1P_PROFILEDATA :
STRUCT
	ALRPROFILEPOS : ARRAY [1..8] OF LREAL;
	ALRPROFILEVEL : ARRAY [1..8] OF LREAL;
	ALRPROFILEACC : ARRAY [1..8] OF LREAL;
	ALRPROFILETIME : ARRAY [1..8] OF LREAL;
	ALRPROFILEJERK : ARRAY [1..8] OF LREAL;
END_STRUCT
END_TYPE

(* ---- L_MB1P_PROFILEPARAMETER.dut ---- *)
TYPE L_MB1P_PROFILEPARAMETER :
STRUCT
	LRTARGETPOS : LREAL;
	LRTARGETVEL : LREAL;
	LRTARGETACC : LREAL;
	LRMAXVEL : LREAL;
	LRMAXACC : LREAL;
	LRMAXDEC : LREAL;
	LRJERKACC : LREAL;
	LRJERKDEC : LREAL;
END_STRUCT
END_TYPE

(* ---- L_MB1P_PROFILEPHASEDATA.dut ---- *)
TYPE L_MB1P_PROFILEPHASEDATA :
STRUCT
	T : LREAL;
	DV : LREAL;
	DS : LREAL;
END_STRUCT
END_TYPE

(* ---- L_MB1P_PROFILETYPE.dut ---- *)
TYPE L_MB1P_PROFILETYPE :
(
	POLY_4TH_ORDER := 0,
	POLY_2TH_ORDER := 1,
	POLY_5TH_ORDER := 2
);
END_TYPE

(* ---- L_MB1P_SCALINGMODE.dut ---- *)
TYPE L_MB1P_SCALINGMODE :
(
	X_ZERO := 0,
	ABSOLUTE := 1,
	RELATIVE := 2
);
END_TYPE

(* ---- L_MB1P_SCXYZCPROFILE.dut ---- *)
TYPE L_MB1P_SCXYZCPROFILE :
STRUCT
	LRXPOS : LREAL;
	LRYPOS : LREAL;
	LRZPOS : LREAL;
	LRCPOS : LREAL;
	LRPATHVEL : LREAL := 10;
	LRPATHACC : LREAL := 100;
	LRPATHDEC : LREAL := 100;
	LRBLENDINGRADIUS : LREAL;
	XHALT : BOOL;
END_STRUCT
END_TYPE

(* ---- L_MB1P_STATES.dut ---- *)
TYPE L_MB1P_STATES :
(
	INIT := 1,
	READY := 2,
	HOMING := 3,
	JOGGING := 10,
	JOGPOS := 11,
	JOGNEG := 12,
	POSITION_TRIMMING := 20,
	TRIM_POS_PLUS := 21,
	TRIM_POS_MINUS := 22,
	SYNCPOS := 30,
	POS_IS_SYNCHRONISED := 31,
	POSITIONING_TO_START_POS := 32,
	SYNCSPEED := 40,
	SPEED_IS_SYNCHRONISED := 41,
	DECOUPLED_LOCAL_DRIVING := 50,
	CONTMOTION := 60,
	PREPARING_PATH := 61,
	CHECK_LIMITS := 62,
	SYNCLINEVEL := 70,
	CAMMING := 80,
	CAMMING_DONE := 81,
	CLUTCH_OPEN_INSTANT := 82,
	CLUTCH_CLOSE := 83,
	CLUTCH_OPEN := 84,
	CYCLICMOTION := 130,
	SETPARAMETERS := 140,
	CAMSEQUENCER_LOADCAMTABLE := 150,
	CAMSEQUENCER_CYCLICCAM1 := 151,
	CAMSEQUENCER_CYCLICCAM3 := 152,
	CAMSEQUENCER_CAM1CYCLICCAM3CAM1 := 153,
	CAMSEQUENCER_CAM1CAM2CYCLICCAM3CAM4CAM1 := 154,
	CALCULATION := 798,
	BUSY := 799,
	DONE := 800,
	EMERGENCYSTOP := 991,
	SLOWSTOP := 992,
	ABC := 993,
	STANDBY := 994,
	HALT := 995,
	STOP := 996,
	QUICKSTOP := 997,
	SERVICE := 998,
	ERROR := 999,
	SYSTEMFAULT := 1000
);
END_TYPE

(* ---- L_TF1P_CAMSEQUENCEMODE.dut ---- *)
TYPE L_TF1P_CAMSEQUENCEMODE :
(
	CYCLICCAM1 := 0,
	CYCLICCAM3 := 1,
	CAM1_CYCLICCAM3_CAM1 := 2,
	CAM1_CAM2_CYCLICCAM3_CAM4_CAM1 := 3
);
END_TYPE

(* ---- L_TF1P_CAMTABLE.dut ---- *)
TYPE L_TF1P_CAMTABLE :
(
	NOCAMTABLE := 0,
	CAMTABLE1 := 1,
	CAMTABLE2 := 2,
	CAMTABLE3 := 3,
	CAMTABLE4 := 4
);
END_TYPE

(* ---- L_TF1P_DIRECTION.dut ---- *)
TYPE L_TF1P_DIRECTION :
(
	BOTH := 0,
	DIRECTIONMASTER := 1
);
END_TYPE

(* ---- L_TF1P_OFFSETMODE.dut ---- *)
TYPE L_TF1P_OFFSETMODE :
(
	X_ZERO := 0,
	DIRECT := 1,
	RAMP_IN := 2,
	DIRECT_BEFOR_SCALE := 3,
	RAMP_IN_BEFOR_SCALE := 4
);
END_TYPE

(* ---- L_TF1P_PROFILETYPE.dut ---- *)
TYPE L_TF1P_PROFILETYPE :
(
	POLY_4TH_ORDER := 0,
	POLY_2TH_ORDER := 1,
	POLY_5TH_ORDER := 2
);
END_TYPE

(* ---- L_TF1P_SCALINGMODE.dut ---- *)
TYPE L_TF1P_SCALINGMODE :
(
	X_ZERO := 0,
	ABSOLUTE := 1,
	RELATIVE := 2,
	RAMP_ABSOLUTE := 3,
	RAMP_RELATIVE := 4
);
END_TYPE

(* ---- L_TF1P_STATES.dut ---- *)
TYPE L_TF1P_STATES :
(
	INIT := 1,
	READY := 2,
	HOMING := 3,
	JOGGING := 10,
	JOGPOS := 11,
	JOGNEG := 12,
	POSITION_TRIMMING := 20,
	TRIM_POS_PLUS := 21,
	TRIM_POS_MINUS := 22,
	SYNCPOS := 30,
	POS_IS_SYNCHRONISED := 31,
	POSITIONING_TO_START_POS := 32,
	SYNCSPEED := 40,
	SPEED_IS_SYNCHRONISED := 41,
	DECOUPLED_LOCAL_DRIVING := 50,
	CONTMOTION := 60,
	PREPARING_PATH := 61,
	CHECK_LIMITS := 62,
	SYNCLINEVEL := 70,
	CAMMING := 80,
	CAMMING_DONE := 81,
	CLUTCH_OPEN_INSTANT := 82,
	CLUTCH_CLOSE := 83,
	CLUTCH_OPEN := 84,
	CYCLICMOTION := 130,
	SETPARAMETERS := 140,
	CAMSEQUENCER_LOADCAMTABLE := 150,
	CAMSEQUENCER_CYCLICCAM1 := 151,
	CAMSEQUENCER_CYCLICCAM3 := 152,
	CAMSEQUENCER_CAM1CYCLICCAM3CAM1 := 153,
	CAMSEQUENCER_CAM1CAM2CYCLICCAM3CAM4CAM1 := 154,
	STANDBY := 994,
	HALT := 995,
	STOP := 996,
	QUICKSTOP := 997,
	SERVICE := 998,
	ERROR := 999
);
END_TYPE

(* ---- L_TF1P_SYNCDIRECTION.dut ---- *)
TYPE L_TF1P_SYNCDIRECTION :
(
	MCNEGATIVEDIRECTION := -1,
	MCCURRENTDIRECTION := 0,
	MCPOSITIVEDIRECTION := 1,
	MCSHORTESTWAY := 2
);
END_TYPE

(* ---- L_TF1P_SYNCMODE.dut ---- *)
TYPE L_TF1P_SYNCMODE :
(
	ABSOLUTE := 0,
	RELATIVE := 1,
	RAMP_TIME := 3,
	RAMP_VELACC := 4,
	RAMP_DIST := 5,
	RAMP_RELATIVE := 7
);
END_TYPE

(* ---- L_TF1P_TPMODE.dut ---- *)
TYPE L_TF1P_TPMODE :
(
	TPFROMMASTER := 0,
	TPFROMSLAVE := 1,
	TPFROMEXTERNAL := 2
);
END_TYPE

(* ---- L_TF1P_TRIMMODE.dut ---- *)
TYPE L_TF1P_TRIMMODE :
(
	VELOCITY := 0,
	POSITION := 1
);
END_TYPE

(* ---- L_TT1P_ADAPTSPDCTRLGAINMODE.dut ---- *)
TYPE L_TT1P_ADAPTSPDCTRLGAINMODE :
(
	DIAMTOSQUARE := 0,
	DIAM := 1,
	INERTIA := 2
);
END_TYPE

(* ---- L_TT1P_CAMDATAXYVA.dut ---- *)
TYPE L_TT1P_CAMDATAXYVA :
STRUCT
	LRX : LREAL;
	LRY : LREAL;
	LRYS : LREAL;
	LRYSS : LREAL;
	LRYSSS : LREAL;
END_STRUCT
END_TYPE

(* ---- L_TT1P_CAMSEQUENCEMODE.dut ---- *)
TYPE L_TT1P_CAMSEQUENCEMODE :
(
	CYCLICCAM1 := 0,
	CYCLICCAM3 := 1,
	CAM1_CYCLICCAM3_CAM1 := 2,
	CAM1_CAM2_CYCLICCAM3_CAM4_CAM1 := 3
);
END_TYPE

(* ---- L_TT1P_CAMTABLE.dut ---- *)
TYPE L_TT1P_CAMTABLE :
(
	NOCAMTABLE := 0,
	CAMTABLE1 := 1,
	CAMTABLE2 := 2,
	CAMTABLE3 := 3,
	CAMTABLE4 := 4
);
END_TYPE

(* ---- L_TT1P_CUTTINGMODEBASE.dut ---- *)
TYPE L_TT1P_CUTTINGMODEBASE :
(
	CUT_LENGTH := 0,
	FLOW_PACKER := 1
);
END_TYPE

(* ---- L_TT1P_CUTTINGMODESTATE.dut ---- *)
TYPE L_TT1P_CUTTINGMODESTATE :
(
	CUT_LENGTH := 0,
	FLOW_PACKER := 1,
	CUT_LENGTH_TP_CORRECTION := 2,
	CUT_ON_TP := 3
);
END_TYPE

(* ---- L_TT1P_DANCERCTRLSTOPMODE.dut ---- *)
TYPE L_TT1P_DANCERCTRLSTOPMODE :
(
	HALT := 0,
	MOVEABS := 1,
	MOVEREL := 2,
	MOVEABSSHORTESTWAY := 3
);
END_TYPE

(* ---- L_TT1P_DANCERLIMITMODE.dut ---- *)
TYPE L_TT1P_DANCERLIMITMODE :
(
	AUTOMATIC := 0,
	SCPARDANCERLIMITS := 1,
	TEACHEDDANCERLIMITS := 2
);
END_TYPE

(* ---- L_TT1P_DIRECTION.dut ---- *)
TYPE L_TT1P_DIRECTION :
(
	BOTH := 0,
	DIRECTIONMASTER := 1
);
END_TYPE

(* ---- L_TT1P_EMODESFLYINGSAW.dut ---- *)
TYPE L_TT1P_EMODESFLYINGSAW :
(
	LENGTHCONTROLLED := 0,
	MARKCONTROLLED := 1
);
END_TYPE

(* ---- L_TT1P_MOVEABSPROFILEDATA.dut ---- *)
TYPE L_TT1P_MOVEABSPROFILEDATA :
STRUCT
	LRPOS_DIST : LREAL;
	LRVEL : LREAL := 0;
	LRACC : LREAL := 0;
	LRDEC : LREAL := 0;
	LRJERKACC : LREAL := 0;
	LRJERKDEC : LREAL := 0;
END_STRUCT
END_TYPE

(* ---- L_TT1P_OFFSETMODE.dut ---- *)
TYPE L_TT1P_OFFSETMODE :
(
	X_ZERO := 0,
	DIRECT := 1,
	RAMP_IN := 2
);
END_TYPE

(* ---- L_TT1P_OFFSETMODESLAVE.dut ---- *)
TYPE L_TT1P_OFFSETMODESLAVE :
(
	X_ZERO := 0,
	DIRECT := 1,
	RAMP_IN := 2,
	DIRECT_BEFOR_SCALE := 3,
	RAMP_IN_BEFOR_SCALE := 4
);
END_TYPE

(* ---- L_TT1P_OSCILLATIONCOMPENSATIONDATA.dut ---- *)
TYPE L_TT1P_OSCILLATIONCOMPENSATIONDATA :
STRUCT
	XVALID : BOOL;
	LRPOSSCALED : LREAL;
	LRLOADSCALED : LREAL;
	LREINGENFREQUENCY : LREAL;
	LRAMPRATION : LREAL;
END_STRUCT
END_TYPE

(* ---- L_TT1P_PERSISTENTVARWINDER.dut ---- *)
TYPE L_TT1P_PERSISTENTVARWINDER :
STRUCT
	LRDIAM : LREAL;
	LRMATERIALCOUNTER : LREAL;
	LIREVCOUNTER : LINT;
	LRREVCOUNTERRESIDUAL : LREAL;
	XUPPERPOSTEACHED : BOOL;
	XLOWERPOSTEACHED : BOOL;
	LRDANCERUPPERLIMIT : LREAL;
	LRDANCERLOWERLIMIT : LREAL;
END_STRUCT
END_TYPE

(* ---- L_TT1P_PICKANDPLACEPATHMODE.dut ---- *)
TYPE L_TT1P_PICKANDPLACEPATHMODE :
(
	LINEAR := 0,
	ELLIPTICAL := 1
);
END_TYPE

(* ---- L_TT1P_POSITIONINGMODE.dut ---- *)
TYPE L_TT1P_POSITIONINGMODE :
(
	ABSOLUTE := 0,
	ABSOLUTE_TP := 1,
	RELATIVE := 2,
	RELATIVE_TP := 3,
	VELOCITY := 4,
	VELOCITY_TP := 5,
	ABSOLUTE_CW_MODULO := 6,
	ABSOLUTE_CW_MODULO_TP := 7,
	ABSOLUTE_CCW_MODULO := 8,
	ABSOLUTE_CCW_MODULO_TP := 9,
	ABSOLUTE_SHORTEST_WAY := 10,
	ABSOLUTE_SHORTEST_WAY_TP := 11
);
END_TYPE

(* ---- L_TT1P_POSITIONPROFILE.dut ---- *)
TYPE L_TT1P_POSITIONPROFILE :
STRUCT
	EPOSITIONINGMODE : L_TT1P_PositioningMode := L_TT1P_PositioningMode.relative;
	LRPOSITION : LREAL := 0;
	LRVELOCITY : LREAL := 0;
	LRACCELERATION : LREAL := 0;
	LRDECELERATION : LREAL := 0;
	LRJERK : LREAL := 0;
	LRFINALVELOCITY : LREAL := 0;
	LRTPWINDOWNEG : LREAL := 0;
	LRTPWINDOWPOS : LREAL := 0;
	ETPPROFILE : L_TT1P_ProfileNumber := L_TT1P_ProfileNumber.No_Profile;
	ESEQUENCEPROFILE : L_TT1P_ProfileNumber := L_TT1P_ProfileNumber.No_Profile;
END_STRUCT
END_TYPE

(* ---- L_TT1P_PROFILEGENERATORDATA.dut ---- *)
TYPE L_TT1P_PROFILEGENERATORDATA :
STRUCT
	ALRPROFILETIME : ARRAY [0..8] OF LREAL;
	ALRPROFILEPOS : ARRAY [0..8] OF LREAL;
	ALRPROFILEVEL : ARRAY [0..8] OF LREAL;
	ALRPROFILEACC : ARRAY [0..8] OF LREAL;
	ALRPROFILEJERK : ARRAY [0..8] OF LREAL;
END_STRUCT
END_TYPE

(* ---- L_TT1P_PROFILENUMBER.dut ---- *)
TYPE L_TT1P_PROFILENUMBER :
(
	NO_PROFILE := 0,
	PROFILE_1 := 1,
	PROFILE_2 := 2,
	PROFILE_3 := 3,
	PROFILE_4 := 4,
	PROFILE_5 := 5,
	PROFILE_6 := 6,
	PROFILE_7 := 7,
	PROFILE_8 := 8,
	PROFILE_9 := 9,
	PROFILE_10 := 10,
	PROFILE_11 := 11,
	PROFILE_12 := 12,
	PROFILE_13 := 13,
	PROFILE_14 := 14,
	PROFILE_15 := 15,
	PROFILE_16 := 16
);
END_TYPE

(* ---- L_TT1P_PROFILES.dut ---- *)
TYPE L_TT1P_PROFILES :
STRUCT
	PROFILE : ARRAY [1..16] OF L_TT1P_PositionProfile;
END_STRUCT
END_TYPE

(* ---- L_TT1P_PROFILETYPE.dut ---- *)
TYPE L_TT1P_PROFILETYPE :
(
	POLY_4TH_ORDER := 0,
	POLY_2TH_ORDER := 1,
	POLY_5TH_ORDER := 2
);
END_TYPE

(* ---- L_TT1P_REGULATORONMODE.dut ---- *)
TYPE L_TT1P_REGULATORONMODE :
(
	DIRECTLYFROMINPUT := 0,
	AUTODISABLE := 1
);
END_TYPE

(* ---- L_TT1P_SCALINGMODE.dut ---- *)
TYPE L_TT1P_SCALINGMODE :
(
	X_ZERO := 0,
	ABSOLUTE := 1,
	RELATIVE := 2,
	RAMP_ABSOLUTE := 3,
	RAMP_RELATIVE := 4
);
END_TYPE

(* ---- L_TT1P_SCAP_ELECTRICALSHAFTPOSBASE.dut ---- *)
TYPE L_TT1P_SCAP_ELECTRICALSHAFTPOSBASE :
STRUCT
END_STRUCT
END_TYPE

(* ---- L_TT1P_SCAP_ELECTRICALSHAFTPOSHIGH.dut ---- *)
TYPE L_TT1P_SCAP_ELECTRICALSHAFTPOSHIGH :
STRUCT
END_STRUCT
END_TYPE

(* ---- L_TT1P_SCAP_ELECTRICALSHAFTPOSSTATE.dut ---- *)
TYPE L_TT1P_SCAP_ELECTRICALSHAFTPOSSTATE :
STRUCT
END_STRUCT
END_TYPE

(* ---- L_TT1P_SCAP_ELECTRICALSHAFTVELBASE.dut ---- *)
TYPE L_TT1P_SCAP_ELECTRICALSHAFTVELBASE :
STRUCT
END_STRUCT
END_TYPE

(* ---- L_TT1P_SCAP_ELECTRICALSHAFTVELHIGH.dut ---- *)
TYPE L_TT1P_SCAP_ELECTRICALSHAFTVELHIGH :
STRUCT
END_STRUCT
END_TYPE

(* ---- L_TT1P_SCAP_ELECTRICALSHAFTVELSTATE.dut ---- *)
TYPE L_TT1P_SCAP_ELECTRICALSHAFTVELSTATE :
STRUCT
END_STRUCT
END_TYPE

(* ---- L_TT1P_SCAP_FLEXCAMBASE.dut ---- *)
TYPE L_TT1P_SCAP_FLEXCAMBASE :
STRUCT
END_STRUCT
END_TYPE

(* ---- L_TT1P_SCAP_FLEXCAMSTATE.dut ---- *)
TYPE L_TT1P_SCAP_FLEXCAMSTATE :
STRUCT
END_STRUCT
END_TYPE

(* ---- L_TT1P_SCAP_FLYINGSAWBASE.dut ---- *)
TYPE L_TT1P_SCAP_FLYINGSAWBASE :
STRUCT
END_STRUCT
END_TYPE

(* ---- L_TT1P_SCAP_FLYINGSAWSTATE.dut ---- *)
TYPE L_TT1P_SCAP_FLYINGSAWSTATE :
STRUCT
END_STRUCT
END_TYPE

(* ---- L_TT1P_SCAP_PICKANDPLACEBASE.dut ---- *)
TYPE L_TT1P_SCAP_PICKANDPLACEBASE :
STRUCT
END_STRUCT
END_TYPE

(* ---- L_TT1P_SCAP_PICKANDPLACEHIGH.dut ---- *)
TYPE L_TT1P_SCAP_PICKANDPLACEHIGH :
STRUCT
END_STRUCT
END_TYPE

(* ---- L_TT1P_SCAP_PICKANDPLACESTATE.dut ---- *)
TYPE L_TT1P_SCAP_PICKANDPLACESTATE :
STRUCT
END_STRUCT
END_TYPE

(* ---- L_TT1P_SCAP_REGISTERCONTROLBASE.dut ---- *)
TYPE L_TT1P_SCAP_REGISTERCONTROLBASE :
STRUCT
END_STRUCT
END_TYPE

(* ---- L_TT1P_SCAP_REGISTERCONTROLSTATE.dut ---- *)
TYPE L_TT1P_SCAP_REGISTERCONTROLSTATE :
STRUCT
END_STRUCT
END_TYPE

(* ---- L_TT1P_SCAP_SMARTTRACKBASE.dut ---- *)
TYPE L_TT1P_SCAP_SMARTTRACKBASE :
STRUCT
END_STRUCT
END_TYPE

(* ---- L_TT1P_SCAP_SMARTTRACKSTATE.dut ---- *)
TYPE L_TT1P_SCAP_SMARTTRACKSTATE :
STRUCT
END_STRUCT
END_TYPE

(* ---- L_TT1P_SCAP_STACKERCRANEAXISCONTROLBASE.dut ---- *)
TYPE L_TT1P_SCAP_STACKERCRANEAXISCONTROLBASE :
STRUCT
END_STRUCT
END_TYPE

(* ---- L_TT1P_SCAP_STACKERCRANEHEADCONTROLBASE.dut ---- *)
TYPE L_TT1P_SCAP_STACKERCRANEHEADCONTROLBASE :
STRUCT
END_STRUCT
END_TYPE

(* ---- L_TT1P_SCAP_TABLEPOSITIONINGBASE.dut ---- *)
TYPE L_TT1P_SCAP_TABLEPOSITIONINGBASE :
STRUCT
END_STRUCT
END_TYPE

(* ---- L_TT1P_SCAP_TM_CROSSCUTTERBASE.dut ---- *)
TYPE L_TT1P_SCAP_TM_CROSSCUTTERBASE :
STRUCT
END_STRUCT
END_TYPE

(* ---- L_TT1P_SCAP_TM_CROSSCUTTERHIGH.dut ---- *)
TYPE L_TT1P_SCAP_TM_CROSSCUTTERHIGH :
STRUCT
END_STRUCT
END_TYPE

(* ---- L_TT1P_SCAP_TM_CROSSCUTTERSTATE.dut ---- *)
TYPE L_TT1P_SCAP_TM_CROSSCUTTERSTATE :
STRUCT
END_STRUCT
END_TYPE

(* ---- L_TT1P_SCAP_WINDERDANCERCTRLBASE.dut ---- *)
TYPE L_TT1P_SCAP_WINDERDANCERCTRLBASE :
STRUCT
END_STRUCT
END_TYPE

(* ---- L_TT1P_SCAP_WINDERDANCERCTRLHIGH.dut ---- *)
TYPE L_TT1P_SCAP_WINDERDANCERCTRLHIGH :
STRUCT
END_STRUCT
END_TYPE

(* ---- L_TT1P_SCAP_WINDERDANCERCTRLSTATE.dut ---- *)
TYPE L_TT1P_SCAP_WINDERDANCERCTRLSTATE :
STRUCT
END_STRUCT
END_TYPE

(* ---- L_TT1P_SCAP_WINDERTENSIONCTRLBASE.dut ---- *)
TYPE L_TT1P_SCAP_WINDERTENSIONCTRLBASE :
STRUCT
END_STRUCT
END_TYPE

(* ---- L_TT1P_SCAP_WINDERTENSIONCTRLHIGH.dut ---- *)
TYPE L_TT1P_SCAP_WINDERTENSIONCTRLHIGH :
STRUCT
END_STRUCT
END_TYPE

(* ---- L_TT1P_SCAP_WINDERTENSIONCTRLSTATE.dut ---- *)
TYPE L_TT1P_SCAP_WINDERTENSIONCTRLSTATE :
STRUCT
END_STRUCT
END_TYPE

(* ---- L_TT1P_SCCOM_STACKERCRANEDATABUS.dut ---- *)
TYPE L_TT1P_SCCOM_STACKERCRANEDATABUS :
STRUCT
END_STRUCT
END_TYPE

(* ---- L_TT1P_SCERRORINFO.dut ---- *)
TYPE L_TT1P_SCERRORINFO :
STRUCT
	XERROR : BOOL;
	XWARNING : BOOL;
	EERRORID : L_IE1P_Error;
	XAXISERROR : BOOL;
	XAXISWARNING : BOOL;
	EAXISERRORID : L_IE1P_Error;
	XDRIVEERROR : BOOL;
	XDRIVEWARNING : BOOL;
	DWDRIVEERRORID : DWORD;
END_STRUCT
END_TYPE

(* ---- L_TT1P_SCPAR_BASICMOTIONBASE.dut ---- *)
TYPE L_TT1P_SCPAR_BASICMOTIONBASE :
STRUCT
END_STRUCT
END_TYPE

(* ---- L_TT1P_SCPAR_CROSSCUTTERBASE.dut ---- *)
TYPE L_TT1P_SCPAR_CROSSCUTTERBASE :
STRUCT
END_STRUCT
END_TYPE

(* ---- L_TT1P_SCPAR_CROSSCUTTERSTATE.dut ---- *)
TYPE L_TT1P_SCPAR_CROSSCUTTERSTATE :
STRUCT
END_STRUCT
END_TYPE

(* ---- L_TT1P_SCPAR_ELECTRICALSHAFTPOSBASE.dut ---- *)
TYPE L_TT1P_SCPAR_ELECTRICALSHAFTPOSBASE :
STRUCT
END_STRUCT
END_TYPE

(* ---- L_TT1P_SCPAR_ELECTRICALSHAFTPOSHIGH.dut ---- *)
TYPE L_TT1P_SCPAR_ELECTRICALSHAFTPOSHIGH :
STRUCT
END_STRUCT
END_TYPE

(* ---- L_TT1P_SCPAR_ELECTRICALSHAFTPOSSTATE.dut ---- *)
TYPE L_TT1P_SCPAR_ELECTRICALSHAFTPOSSTATE :
STRUCT
END_STRUCT
END_TYPE

(* ---- L_TT1P_SCPAR_ELECTRICALSHAFTVELBASE.dut ---- *)
TYPE L_TT1P_SCPAR_ELECTRICALSHAFTVELBASE :
STRUCT
END_STRUCT
END_TYPE

(* ---- L_TT1P_SCPAR_ELECTRICALSHAFTVELHIGH.dut ---- *)
TYPE L_TT1P_SCPAR_ELECTRICALSHAFTVELHIGH :
STRUCT
END_STRUCT
END_TYPE

(* ---- L_TT1P_SCPAR_ELECTRICALSHAFTVELSTATE.dut ---- *)
TYPE L_TT1P_SCPAR_ELECTRICALSHAFTVELSTATE :
STRUCT
END_STRUCT
END_TYPE

(* ---- L_TT1P_SCPAR_FLEXCAMBASE.dut ---- *)
TYPE L_TT1P_SCPAR_FLEXCAMBASE :
STRUCT
END_STRUCT
END_TYPE

(* ---- L_TT1P_SCPAR_FLEXCAMSTATE.dut ---- *)
TYPE L_TT1P_SCPAR_FLEXCAMSTATE :
STRUCT
END_STRUCT
END_TYPE

(* ---- L_TT1P_SCPAR_FLYINGSAWBASE.dut ---- *)
TYPE L_TT1P_SCPAR_FLYINGSAWBASE :
STRUCT
END_STRUCT
END_TYPE

(* ---- L_TT1P_SCPAR_FLYINGSAWSTATE.dut ---- *)
TYPE L_TT1P_SCPAR_FLYINGSAWSTATE :
STRUCT
END_STRUCT
END_TYPE

(* ---- L_TT1P_SCPAR_PICKANDPLACEBASE.dut ---- *)
TYPE L_TT1P_SCPAR_PICKANDPLACEBASE :
STRUCT
END_STRUCT
END_TYPE

(* ---- L_TT1P_SCPAR_PICKANDPLACEHIGH.dut ---- *)
TYPE L_TT1P_SCPAR_PICKANDPLACEHIGH :
STRUCT
END_STRUCT
END_TYPE

(* ---- L_TT1P_SCPAR_PICKANDPLACESTATE.dut ---- *)
TYPE L_TT1P_SCPAR_PICKANDPLACESTATE :
STRUCT
END_STRUCT
END_TYPE

(* ---- L_TT1P_SCPAR_REGISTERCONTROLBASE.dut ---- *)
TYPE L_TT1P_SCPAR_REGISTERCONTROLBASE :
STRUCT
END_STRUCT
END_TYPE

(* ---- L_TT1P_SCPAR_REGISTERCONTROLSTATE.dut ---- *)
TYPE L_TT1P_SCPAR_REGISTERCONTROLSTATE :
STRUCT
END_STRUCT
END_TYPE

(* ---- L_TT1P_SCPAR_SMARTTRACKBASE.dut ---- *)
TYPE L_TT1P_SCPAR_SMARTTRACKBASE :
STRUCT
END_STRUCT
END_TYPE

(* ---- L_TT1P_SCPAR_SMARTTRACKSTATE.dut ---- *)
TYPE L_TT1P_SCPAR_SMARTTRACKSTATE :
STRUCT
END_STRUCT
END_TYPE

(* ---- L_TT1P_SCPAR_STACKERCRANEAXISCONTROLBASE.dut ---- *)
TYPE L_TT1P_SCPAR_STACKERCRANEAXISCONTROLBASE :
STRUCT
END_STRUCT
END_TYPE

(* ---- L_TT1P_SCPAR_STACKERCRANEHEADCONTROLBASE.dut ---- *)
TYPE L_TT1P_SCPAR_STACKERCRANEHEADCONTROLBASE :
STRUCT
END_STRUCT
END_TYPE

(* ---- L_TT1P_SCPAR_TABLEPOSITIONINGBASE.dut ---- *)
TYPE L_TT1P_SCPAR_TABLEPOSITIONINGBASE :
STRUCT
END_STRUCT
END_TYPE

(* ---- L_TT1P_SCPAR_VIRTUALMASTERBASE.dut ---- *)
TYPE L_TT1P_SCPAR_VIRTUALMASTERBASE :
STRUCT
END_STRUCT
END_TYPE

(* ---- L_TT1P_SCPAR_VIRTUALMASTERHIGH.dut ---- *)
TYPE L_TT1P_SCPAR_VIRTUALMASTERHIGH :
STRUCT
END_STRUCT
END_TYPE

(* ---- L_TT1P_SCPAR_VIRTUALMASTERSTATE.dut ---- *)
TYPE L_TT1P_SCPAR_VIRTUALMASTERSTATE :
STRUCT
END_STRUCT
END_TYPE

(* ---- L_TT1P_SCPAR_WINDERDANCERCTRLBASE.dut ---- *)
TYPE L_TT1P_SCPAR_WINDERDANCERCTRLBASE :
STRUCT
END_STRUCT
END_TYPE

(* ---- L_TT1P_SCPAR_WINDERDANCERCTRLHIGH.dut ---- *)
TYPE L_TT1P_SCPAR_WINDERDANCERCTRLHIGH :
STRUCT
END_STRUCT
END_TYPE

(* ---- L_TT1P_SCPAR_WINDERDANCERCTRLSTATE.dut ---- *)
TYPE L_TT1P_SCPAR_WINDERDANCERCTRLSTATE :
STRUCT
END_STRUCT
END_TYPE

(* ---- L_TT1P_SCPAR_WINDERTENSIONCTRLBASE.dut ---- *)
TYPE L_TT1P_SCPAR_WINDERTENSIONCTRLBASE :
STRUCT
END_STRUCT
END_TYPE

(* ---- L_TT1P_SCPAR_WINDERTENSIONCTRLHIGH.dut ---- *)
TYPE L_TT1P_SCPAR_WINDERTENSIONCTRLHIGH :
STRUCT
END_STRUCT
END_TYPE

(* ---- L_TT1P_SCPAR_WINDERTENSIONCTRLSTATE.dut ---- *)
TYPE L_TT1P_SCPAR_WINDERTENSIONCTRLSTATE :
STRUCT
END_STRUCT
END_TYPE

(* ---- L_TT1P_SCPROFILEPAR.dut ---- *)
TYPE L_TT1P_SCPROFILEPAR :
STRUCT
END_STRUCT
END_TYPE

(* ---- L_TT1P_SCSF_ELECTRICALSHAFTPOSBASE.dut ---- *)
TYPE L_TT1P_SCSF_ELECTRICALSHAFTPOSBASE :
STRUCT
END_STRUCT
END_TYPE

(* ---- L_TT1P_SCSF_ELECTRICALSHAFTPOSHIGH.dut ---- *)
TYPE L_TT1P_SCSF_ELECTRICALSHAFTPOSHIGH :
STRUCT
END_STRUCT
END_TYPE

(* ---- L_TT1P_SCSF_ELECTRICALSHAFTPOSSTATE.dut ---- *)
TYPE L_TT1P_SCSF_ELECTRICALSHAFTPOSSTATE :
STRUCT
END_STRUCT
END_TYPE

(* ---- L_TT1P_SCSF_ELECTRICALSHAFTVELBASE.dut ---- *)
TYPE L_TT1P_SCSF_ELECTRICALSHAFTVELBASE :
STRUCT
END_STRUCT
END_TYPE

(* ---- L_TT1P_SCSF_ELECTRICALSHAFTVELHIGH.dut ---- *)
TYPE L_TT1P_SCSF_ELECTRICALSHAFTVELHIGH :
STRUCT
END_STRUCT
END_TYPE

(* ---- L_TT1P_SCSF_ELECTRICALSHAFTVELSTATE.dut ---- *)
TYPE L_TT1P_SCSF_ELECTRICALSHAFTVELSTATE :
STRUCT
END_STRUCT
END_TYPE

(* ---- L_TT1P_SCSF_FLEXCAMBASE.dut ---- *)
TYPE L_TT1P_SCSF_FLEXCAMBASE :
STRUCT
END_STRUCT
END_TYPE

(* ---- L_TT1P_SCSF_FLEXCAMSTATE.dut ---- *)
TYPE L_TT1P_SCSF_FLEXCAMSTATE :
STRUCT
END_STRUCT
END_TYPE

(* ---- L_TT1P_SCSF_FLYINGSAWBASE.dut ---- *)
TYPE L_TT1P_SCSF_FLYINGSAWBASE :
STRUCT
END_STRUCT
END_TYPE

(* ---- L_TT1P_SCSF_FLYINGSAWSTATE.dut ---- *)
TYPE L_TT1P_SCSF_FLYINGSAWSTATE :
STRUCT
END_STRUCT
END_TYPE

(* ---- L_TT1P_SCSF_PICKANDPLACEBASE.dut ---- *)
TYPE L_TT1P_SCSF_PICKANDPLACEBASE :
STRUCT
END_STRUCT
END_TYPE

(* ---- L_TT1P_SCSF_PICKANDPLACEHIGH.dut ---- *)
TYPE L_TT1P_SCSF_PICKANDPLACEHIGH :
STRUCT
END_STRUCT
END_TYPE

(* ---- L_TT1P_SCSF_PICKANDPLACESTATE.dut ---- *)
TYPE L_TT1P_SCSF_PICKANDPLACESTATE :
STRUCT
END_STRUCT
END_TYPE

(* ---- L_TT1P_SCSF_REGISTERCONTROLBASE.dut ---- *)
TYPE L_TT1P_SCSF_REGISTERCONTROLBASE :
STRUCT
END_STRUCT
END_TYPE

(* ---- L_TT1P_SCSF_REGISTERCONTROLSTATE.dut ---- *)
TYPE L_TT1P_SCSF_REGISTERCONTROLSTATE :
STRUCT
END_STRUCT
END_TYPE

(* ---- L_TT1P_SCSF_SMARTTRACKBASE.dut ---- *)
TYPE L_TT1P_SCSF_SMARTTRACKBASE :
STRUCT
END_STRUCT
END_TYPE

(* ---- L_TT1P_SCSF_SMARTTRACKSTATE.dut ---- *)
TYPE L_TT1P_SCSF_SMARTTRACKSTATE :
STRUCT
END_STRUCT
END_TYPE

(* ---- L_TT1P_SCSF_STACKERCRANEAXISCONTROLBASE.dut ---- *)
TYPE L_TT1P_SCSF_STACKERCRANEAXISCONTROLBASE :
STRUCT
END_STRUCT
END_TYPE

(* ---- L_TT1P_SCSF_STACKERCRANEHEADCONTROLBASE.dut ---- *)
TYPE L_TT1P_SCSF_STACKERCRANEHEADCONTROLBASE :
STRUCT
END_STRUCT
END_TYPE

(* ---- L_TT1P_SCSF_TABLEPOSITIONINGBASE.dut ---- *)
TYPE L_TT1P_SCSF_TABLEPOSITIONINGBASE :
STRUCT
END_STRUCT
END_TYPE

(* ---- L_TT1P_SCSF_TM_CROSSCUTTERBASE.dut ---- *)
TYPE L_TT1P_SCSF_TM_CROSSCUTTERBASE :
STRUCT
END_STRUCT
END_TYPE

(* ---- L_TT1P_SCSF_TM_CROSSCUTTERHIGH.dut ---- *)
TYPE L_TT1P_SCSF_TM_CROSSCUTTERHIGH :
STRUCT
END_STRUCT
END_TYPE

(* ---- L_TT1P_SCSF_TM_CROSSCUTTERSTATE.dut ---- *)
TYPE L_TT1P_SCSF_TM_CROSSCUTTERSTATE :
STRUCT
END_STRUCT
END_TYPE

(* ---- L_TT1P_SCSF_WINDERDANCERCTRLBASE.dut ---- *)
TYPE L_TT1P_SCSF_WINDERDANCERCTRLBASE :
STRUCT
END_STRUCT
END_TYPE

(* ---- L_TT1P_SCSF_WINDERDANCERCTRLLHIGH.dut ---- *)
TYPE L_TT1P_SCSF_WINDERDANCERCTRLLHIGH :
STRUCT
END_STRUCT
END_TYPE

(* ---- L_TT1P_SCSF_WINDERDANCERCTRLSTATE.dut ---- *)
TYPE L_TT1P_SCSF_WINDERDANCERCTRLSTATE :
STRUCT
END_STRUCT
END_TYPE

(* ---- L_TT1P_SCSF_WINDERTENSIONCTRLBASE.dut ---- *)
TYPE L_TT1P_SCSF_WINDERTENSIONCTRLBASE :
STRUCT
END_STRUCT
END_TYPE

(* ---- L_TT1P_SCSF_WINDERTENSIONCTRLHIGH.dut ---- *)
TYPE L_TT1P_SCSF_WINDERTENSIONCTRLHIGH :
STRUCT
END_STRUCT
END_TYPE

(* ---- L_TT1P_SCSF_WINDERTENSIONCTRLSTATE.dut ---- *)
TYPE L_TT1P_SCSF_WINDERTENSIONCTRLSTATE :
STRUCT
END_STRUCT
END_TYPE

(* ---- L_TT1P_SOURCEFORCORRWINDOW.dut ---- *)
TYPE L_TT1P_SOURCEFORCORRWINDOW :
(
	MASTER := 0,
	REGISTER := 1,
	SLAVE := 2
);
END_TYPE

(* ---- L_TT1P_STACKERCRANEADDRESS.dut ---- *)
TYPE L_TT1P_STACKERCRANEADDRESS :
(
	HEADCONTROL := 10,
	X_AXIS := 20,
	Y_AXIS := 21,
	AP_AXIS := 31,
	X_SLAVEAXIS1 := 32,
	Y_SLAVEAXIS1 := 33
);
END_TYPE

(* ---- L_TT1P_STATES.dut ---- *)
TYPE L_TT1P_STATES :
(
	INIT := 1,
	READY := 2,
	HOMING := 3,
	JOGGING := 10,
	JOGPOS := 11,
	JOGNEG := 12,
	MOVEVEL := 13,
	MOVEABS := 14,
	MOVEREL := 15,
	EXTERNAL := 17,
	POSITION_TRIMMING := 20,
	TRIM_POS_PLUS := 21,
	TRIM_POS_MINUS := 22,
	SYNCHRONISING_POS := 30,
	POS_IS_SYNCHRONISED := 31,
	POSITIONING_TO_START_POS := 32,
	CAMMING := 33,
	POSITIONING_TO_TARGET_POS := 34,
	POSITIONING_TO_PARK_POS := 35,
	MOVE_TO_TARGET_POS := 36,
	POSITIONING := 38,
	SYNCHRONISING_VEL := 40,
	VEL_IS_SYNCHRONISED := 41,
	DECOUPLED_LOCAL_DRIVING := 50,
	GROUNDSPEED := 51,
	ACC_DEC := 52,
	CONTMOTION := 60,
	SYNCLINEVEL := 70,
	IDENTMINERTIA := 80,
	IDENTDIAMETER := 81,
	IDENTFRICTION := 90,
	DANCERCTRL := 100,
	TENSIONCTRL := 110,
	PREPARING_PATH := 112,
	MOVE_PP := 114,
	CHECK_LIMITS := 115,
	TRANSFORMATION := 116,
	PATH_INTERRUPT := 117,
	SELECTMODEVL := 120,
	SELECTMODECSV := 121,
	SELECTMODECST := 122,
	SELECTMODECSP := 123,
	CYCLICMOTION := 130,
	SETPARAMETERS := 140,
	JOGGING_X := 150,
	JOGGING_Y := 151,
	JOGGING_Z := 152,
	JOGGING_A := 153,
	JOGGING_B := 154,
	JOGGING_C := 155,
	JOGGING_A1 := 156,
	JOGGING_A2 := 157,
	JOGGING_A3 := 158,
	JOGGING_A4 := 159,
	JOGGING_A5 := 160,
	JOGGING_A6 := 161,
	JOGGING_AUX1 := 162,
	JOGGING_AUX2 := 163,
	JOGGING_AUX3 := 164,
	JOGGING_AUX4 := 165,
	JOGGING_AUX5 := 166,
	JOGGING_AUX6 := 167,
	CUTTING := 170,
	IN_PARK_POS := 171,
	ASYNC_PHASE := 172,
	ENTRY_IN_SYNC_PAHSE := 173,
	EXIT_SYNC_PHASE := 175,
	HOLD_IN_PARK_POS := 176,
	CLUTCH_CLOSE := 177,
	CLUTCH_OPEN := 178,
	WAIT_OF_NEXT_CUT := 179,
	STOP_IN_PARK_POS := 180,
	MOVE_TO_INFEED := 181,
	IN_INFEED := 182,
	MOVE_TO_OUTFEED := 183,
	IN_OUTFEED := 184,
	MAGICTRACK := 185,
	MOVE_XY := 186,
	MAINTENANCE := 187,
	BRAKE_TEST := 188,
	BRAKE_GRINDIN := 189,
	TRAVERSING := 190,
	SAW_IN_PROCESS := 200,
	MOVE_TO_PARK_POS := 210,
	DONE := 800,
	EMERGENCYSTOP := 991,
	SLOWSTOP := 992,
	ABC := 993,
	STANDBY := 994,
	STOP := 996,
	QUICKSTOP := 997,
	SERVICE := 998,
	ERROR := 999,
	SYSTEMFAULT := 1000
);
END_TYPE

(* ---- L_TT1P_SYNCDIRECTION.dut ---- *)
TYPE L_TT1P_SYNCDIRECTION :
(
	MCNEGATIVEDIRECTION := -1,
	MCCURRENTDIRECTION := 0,
	MCPOSITIVEDIRECTION := 1
);
END_TYPE

(* ---- L_TT1P_SYNCDIRECTIONELECTRICALSHAFTPOS.dut ---- *)
TYPE L_TT1P_SYNCDIRECTIONELECTRICALSHAFTPOS :
(
	MCNEGATIVEDIRECTION := -1,
	MCPOSITIVEDIRECTION := 1,
	MCSHORTESTWAY := 2
);
END_TYPE

(* ---- L_TT1P_SYNCDIRECTIONVIRTUALMASTER.dut ---- *)
TYPE L_TT1P_SYNCDIRECTIONVIRTUALMASTER :
(
	MCNEGATIVEDIRECTION := -1,
	MCPOSITIVEDIRECTION := 1,
	MCSHORTESTWAY := 2
);
END_TYPE

(* ---- L_TT1P_SYNCMODE.dut ---- *)
TYPE L_TT1P_SYNCMODE :
(
	ABSOLUTE := 0,
	RELATIVE := 1,
	RAMP_POS := 2,
	RAMP_TIME := 3,
	RAMP_VELACC := 4
);
END_TYPE

(* ---- L_TT1P_SYNCMODECROSSCUTTER.dut ---- *)
TYPE L_TT1P_SYNCMODECROSSCUTTER :
(
	CAM_IN := 0,
	POSITIONING := 1
);
END_TYPE

(* ---- L_TT1P_SYNCMODEELECTRICALSHAFTPOS.dut ---- *)
TYPE L_TT1P_SYNCMODEELECTRICALSHAFTPOS :
(
	RAMP_TIME := 3,
	RAMP_VELACC := 4,
	RAMP_DIST := 5
);
END_TYPE

(* ---- L_TT1P_SYNCMODEVIRTUALMASTER.dut ---- *)
TYPE L_TT1P_SYNCMODEVIRTUALMASTER :
(
	RAMP_TIME := 3,
	RAMP_VELACC := 4,
	RAMP_DIST := 5
);
END_TYPE

(* ---- L_TT1P_TENSIONCTRLSTOPMODE.dut ---- *)
TYPE L_TT1P_TENSIONCTRLSTOPMODE :
(
	HALT := 0,
	MOVEABS := 1,
	MOVEREL := 2,
	MOVEABSSHORTESTWAY := 3
);
END_TYPE

(* ---- L_TT1P_TPMODE.dut ---- *)
TYPE L_TT1P_TPMODE :
(
	TPFROMMASTER := 0,
	TPFROMSLAVE := 1,
	TPFROMEXTERNAL := 2
);
END_TYPE

(* ---- L_TT1P_TPMODESINGLEAXIS.dut ---- *)
TYPE L_TT1P_TPMODESINGLEAXIS :
(
	TPFROMTMAXIS := 0,
	TPFROMEXTERNAL := 1
);
END_TYPE

(* ---- L_TT1P_TRACKPICKANDPLACEMODE.dut ---- *)
TYPE L_TT1P_TRACKPICKANDPLACEMODE :
(
	SETTARGET := 0,
	TARGETPOSTOCV1 := 1,
	CV1TOTARGETPOS := 2,
	CV1TOCV2 := 3,
	CV2TOCV1 := 4
);
END_TYPE

(* ---- L_TT1P_TRACKPICKANDPLACETARGET.dut ---- *)
TYPE L_TT1P_TRACKPICKANDPLACETARGET :
(
	MOVEPICKANDPLACEPROFIL := 0,
	SYNCCONVEYOR1 := 1,
	SYNCCONVEYOR2 := 2,
	SYNCCONVEYOR3 := 3,
	SYNCCONVEYOR4 := 4,
	SYNCCONVEYOR5 := 5,
	SYNCCONVEYOR6 := 6,
	SYNCCONVEYOR7 := 7,
	SYNCCONVEYOR8 := 8,
	SYNCCONVEYOR9 := 9,
	SYNCCONVEYOR10 := 10,
	SYNCCONVEYOR11 := 11,
	SYNCCONVEYOR12 := 12,
	SYNCCONVEYOR13 := 13,
	SYNCCONVEYOR14 := 14,
	SYNCCONVEYOR15 := 15,
	SYNCCONVEYOR16 := 16
);
END_TYPE

(* ---- L_TT1P_TRACKPICKANDPLACETARGETSTATUS.dut ---- *)
TYPE L_TT1P_TRACKPICKANDPLACETARGETSTATUS :
(
	INACTIVE := 0,
	MOVETOPARKPOS := 1,
	INPARKPOS := 2,
	MOVETOTARGET := 3,
	INTARGET := 4,
	MOVEFROMTARGET := 5
);
END_TYPE

(* ---- L_TT1P_TRIMMODE.dut ---- *)
TYPE L_TT1P_TRIMMODE :
(
	VELOCITY := 0,
	POSITION := 1
);
END_TYPE

(* ---- L_TT1P_XYBUFFERDATA.dut ---- *)
TYPE L_TT1P_XYBUFFERDATA :
STRUCT
	LRBUFFERPOSITIONPOS : LREAL;
	LRBUFFERPOSITIONNEG : LREAL;
	LRBUFFERVELPOS : LREAL;
	LRBUFFERVELNEG : LREAL;
END_STRUCT
END_TYPE

(* ---- L_TT1P_XYLIMITS.dut ---- *)
TYPE L_TT1P_XYLIMITS :
STRUCT
	LRVELOCITY : LREAL;
	LRACCELERATION : LREAL;
	LRDECELERATION : LREAL;
END_STRUCT
END_TYPE

(* ---- L_TT1P_XYMODE.dut ---- *)
TYPE L_TT1P_XYMODE :
(
	NOTCOORDINATED := 0,
	SYNCSTARTSTOP := 1,
	ASYNCSTARTSYNCSTOP := 2,
	ASYNCSTARTORSTOP := 3,
	ASYNCSTARTSYNCSTOPTIMEOPT := 4,
	ASYNCSTARTORSTOPTIMEOPT := 5
);
END_TYPE

(* ---- L_TT1P_XYPROFILEDATA.dut ---- *)
TYPE L_TT1P_XYPROFILEDATA :
STRUCT
	EPROFILEMODE : L_TT1P_XYProfileMode;
	LRTARGETPOSITION : LREAL;
	LRVELOCITY : LREAL;
	LRACCELERATION : LREAL;
	LRDECELERATION : LREAL;
	LRJERKACCELERATION : LREAL;
	LRJERKDECELERATION : LREAL;
END_STRUCT
END_TYPE

(* ---- L_TT1P_XYPROFILEMODE.dut ---- *)
TYPE L_TT1P_XYPROFILEMODE :
(
	ABSOLUTE := 0,
	RELATIVE := 2
);
END_TYPE

(* ---- SCCTRL_ABC.dut ---- *)
TYPE SCCTRL_ABC :
STRUCT
	XRESETERROR : BOOL;
	XREGULATORON : BOOL;
	XENABLEPOSITIVE : BOOL := TRUE;
	XENABLENEGATIVE : BOOL := TRUE;
	XJOGGINGPOS : BOOL;
	XJOGGINGNEG : BOOL;
	LRJOGGINGSETVEL : LREAL := 100;
	LRJOGGINGSETACC : LREAL := 100;
	LRJOGGINGSETDEC : LREAL := 100;
	LRJOGGINGSETJERK : LREAL := 0;
	XCONTINUOUSUPDATE : BOOL;
	XSTOP : BOOL;
	XHALT : BOOL;
	XMOVEVELEXECUTE : BOOL;
	XMOVEABSEXECUTE : BOOL;
	XMOVERELEXECUTE : BOOL;
	LRSETPOS_DIST : LREAL := 0;
	LRSETVEL : LREAL := 100;
	LRSETACC : LREAL := 100;
	LRSETDEC : LREAL := 100;
	LRSETJERK : LREAL := 0;
	ESETDIRECTION : MC_DIRECTION := MC_DIRECTION.mcPositiveDirection;
	XHOMEEXECUTE : BOOL;
	LRHOMEPOSITION : LREAL := 0;
	XUSEHOMEEXTPARAMETER : BOOL;
	SCHOMEEXTPARAMETER : L_MC1P_HomeParameter;
	SCHOMEEXTTP : MC_TRIGGER_REF;
	XHOMEABSSWITCH : BOOL;
	LROVERRIDEJERK : LREAL := 1;
	LROVERRIDEACC : LREAL := 1;
	LROVERRIDE : LREAL := 1;
END_STRUCT
END_TYPE

(* ---- SCCTRL_AGBC.dut ---- *)
TYPE SCCTRL_AGBC :
STRUCT
	XREGULATORONALL : BOOL;
	XENABLEAXESGROUP : BOOL;
	XRESETAXESGROUP : BOOL;
	LROVERRIDE : LREAL := 1;
	XSTOPALL : BOOL;
	SCPAR : L_MC4P_AGBC_Parameter;
	ECOORDSYSTEM : L_MC4P_CoordSystem := 0;
	XGROUPSTOPEXECUTE : BOOL;
	XMOVEDIRABSEXECUTE : BOOL;
	XMOVEDIRRELEXECUTE : BOOL;
	XMOVELINABSEXECUTE : BOOL;
	XMOVELINRELEXECUTE : BOOL;
	ALRSETPOSDIST : ARRAY [1..12] OF LREAL;
	XGROUPSETPOSEXECUTE : BOOL;
	XGROUPHOMEEXECUTE : BOOL;
	AXHOMEABSSWITCH : ARRAY [1..12] OF BOOL;
	ASCHOMEEXTTP : ARRAY [1..12] OF MC_TRIGGER_REF;
	AXJOGPOS : ARRAY [1..12] OF BOOL;
	AXJOGNEG : ARRAY [1..12] OF BOOL;
	AXMOVEABS : ARRAY [1..12] OF BOOL;
	AXMOVEREL : ARRAY [1..12] OF BOOL;
	ASCCTRLABC : ARRAY [1..18] OF L_MC1P_CtrlABC;
END_STRUCT
END_TYPE

(* ---- SCSTATUS_ABC.dut ---- *)
TYPE SCSTATUS_ABC :
STRUCT
	XINTERNALCONTROLACTIVE : BOOL;
	XERROR : BOOL;
	EERRORID : L_IE1P_Error;
	XFUNBUSY : BOOL;
	XFUNDONE : BOOL;
	XFUNCOMMANDABORTED : BOOL;
	EFUNSTATEACT : L_MC1P_ABC_State;
	ECONTROLMODE : L_MC1P_ControlMode;
	XISHOMED : BOOL;
	XHWLIMITSWITCHNEG : BOOL;
	XHWLIMITSWITCHPOS : BOOL;
	XSWLIMITENABLED : BOOL;
	XSWLIMITSWITCHNEG : BOOL;
	XSWLIMITSWITCHPOS : BOOL;
	EAXISTYPE : L_MC1P_DriveType;
	EAXISSTATE : L_MC1P_AXIS_STATE;
	XAXISREADY : BOOL;
	XAXISENABLED : BOOL;
	XAXISWARNING : BOOL;
	XAXISERROR : BOOL;
	EAXISERRORID : L_IE1P_Error;
	XDRIVEWARNING : BOOL;
	XDRIVEERROR : BOOL;
	DWDRIVEERRORID : DWORD;
	LRACTPOS : LREAL;
	LRACTVEL : LREAL;
	LRSETPOSOUT : LREAL;
	LRSETVELOUT : LREAL;
	LRACTFOLLOWINGERROR : LREAL;
	XCONSTANTVELOCITY : BOOL;
	XACCELERATING : BOOL;
	XDECELERATING : BOOL;
	XDIRECTIONPOSITIVE : BOOL;
	XDIRECTIONNEGATIVE : BOOL;
	XINPOSITION : BOOL;
	XAXISAVAILABLE : BOOL;
	XSTANDSTILLSETVELOCITY : BOOL;
	XSTANDSTILLACTVELOCITY : BOOL;
END_STRUCT
END_TYPE

(* ---- SCSTATUS_AGBC.dut ---- *)
TYPE SCSTATUS_AGBC :
STRUCT
	XINTERNALCONTROLACTIVE : BOOL;
	XERROR : BOOL;
	EERRORID : L_IE1P_Error;
	XFUNBUSY : BOOL;
	XFUNDONE : BOOL;
	XFUNCOMMANDABORTED : BOOL;
	EFUNSTATEACT : L_MC4P_AGBC_State := L_MC4P_AGBC_State.Standby;
	XAXESGROUPHOMED : BOOL;
	XHWLIMITSWITCHANY : BOOL;
	XSWLIMITENABLEDALL : BOOL;
	XSWLIMITSWITCHANY : BOOL;
	EKINEMATICTYPE : L_MC4P_KinematicType;
	EAXESGROUPSTATE : L_MC4P_AxesGroup_State;
	XAXESGROUPENABLED : BOOL;
	XREALAXESREADYALL : BOOL;
	XREALAXESENABLEDALL : BOOL;
	XINPOSITION : BOOL;
	XAXESGROUPWARNING : BOOL;
	XAXESGROUPERROR : BOOL;
	EAXESGROUPERRORID : L_IE1P_Error;
	ALRACTPOS : ARRAY [1..12] OF LREAL;
	ALRACTVEL : ARRAY [1..12] OF LREAL;
	ALRSETPOSOUT : ARRAY [1..12] OF LREAL;
	ALRSETVELOUT : ARRAY [1..12] OF LREAL;
	ALRACTFOLLOWINGERROR : ARRAY [1..12] OF LREAL;
	LRSETPATHVELOUT : LREAL;
	LRSETPATHACCOUT : LREAL;
	LRSETTCPACCOUT : LREAL := 0;
	LRSETROTVELOUT : LREAL := 0;
	LRSETROTACCOUT : LREAL := 0;
	ASCSTATUSABC : ARRAY [1..18] OF L_MC1P_StatusABC;
END_STRUCT
END_TYPE

(* ---- L_MB1P_CONSTANTS.gvl ---- *)
VAR_GLOBAL
	GC_DWCHECKIDTAPPETREF : DWORD := 16#DC34;
	GC_LREPSILON : LREAL := 1E-06;
	GC_POSITIVE_LIMIT_32BIT : LREAL := 2147483647;
	GC_NEGATIVE_LIMIT_32BIT : LREAL := -2147483647;
	GC_PI : LREAL := 3.1415926535897931;
END_VAR

(* ---- L_MB1P_GLOBAL.gvl ---- *)
VAR_GLOBAL
END_VAR

(* ---- ITF_DATABUS.itf ---- *)
INTERFACE ITF_DATABUS
END_INTERFACE

(* ---- ITF_DATABUSPAR.itf ---- *)
INTERFACE ITF_DATABUSPAR
END_INTERFACE

(* ---- ITF_LIST.itf ---- *)
INTERFACE ITF_LIST
END_INTERFACE

(* ---- GETBOOLEANPROPERTY.pou ---- *)
FUNCTION GETBOOLEANPROPERTY : BOOL
VAR_INPUT
	STKEY : WSTRING;
END_VAR
END_FUNCTION

(* ---- GETCOMPANY.pou ---- *)
FUNCTION GETCOMPANY : WSTRING
END_FUNCTION

(* ---- GETNUMBERPROPERTY.pou ---- *)
FUNCTION GETNUMBERPROPERTY : DINT
VAR_INPUT
	STKEY : WSTRING;
END_VAR
END_FUNCTION

(* ---- GETTEXTPROPERTY.pou ---- *)
FUNCTION GETTEXTPROPERTY : WSTRING
VAR_INPUT
	STKEY : WSTRING;
END_VAR
END_FUNCTION

(* ---- GETTEXTPROPERTY2.pou ---- *)
FUNCTION GETTEXTPROPERTY2 : POINTER TO WSTRING
VAR_INPUT
	STKEY : WSTRING;
END_VAR
END_FUNCTION

(* ---- GETTITLE.pou ---- *)
FUNCTION GETTITLE : WSTRING
END_FUNCTION

(* ---- GETVERSION.pou ---- *)
FUNCTION GETVERSION : VERSION
END_FUNCTION

(* ---- GETVERSIONPROPERTY.pou ---- *)
FUNCTION GETVERSIONPROPERTY : VERSION
VAR_INPUT
	STKEY : WSTRING;
END_VAR
END_FUNCTION

(* ---- L_MB1P_CALCDISTBETWEEN3DPOINTS.pou ---- *)
FUNCTION L_MB1P_CALCDISTBETWEEN3DPOINTS : LREAL
VAR_INPUT
	LRX1 : LREAL;
	LRY1 : LREAL;
	LRZ1 : LREAL;
	LRX2 : LREAL;
	LRY2 : LREAL;
	LRZ2 : LREAL;
END_VAR
END_FUNCTION

(* ---- L_MB1P_CALCIDENDIAMETERBASE.pou ---- *)
FUNCTION L_MB1P_CALCIDENDIAMETERBASE : LREAL
VAR_IN_OUT
	LRLINEDIST : LREAL;
	LRDIAMCALCDIST : LREAL;
END_VAR
END_FUNCTION

(* ---- L_MB1P_CALCIDENDIAMETERSTATE.pou ---- *)
FUNCTION L_MB1P_CALCIDENDIAMETERSTATE : LREAL
VAR_IN_OUT
	LRDANCERPOSSTART : LREAL;
	LRDANCERPOSEND : LREAL;
	LRDIAMCALCDIST : LREAL;
	LRDANCERMATERIALLENGTH : LREAL;
END_VAR
END_FUNCTION

(* ---- L_MB1P_CHECK_CAMREFCHANGED.pou ---- *)
FUNCTION L_MB1P_CHECK_CAMREFCHANGED : BOOL
VAR_INPUT
	CAMREFNEW : MC_CAM_REF;
	CAMREFOLD : MC_CAM_REF;
END_VAR
END_FUNCTION

(* ---- L_MB1P_CHECK_CAMREFVALID.pou ---- *)
FUNCTION L_MB1P_CHECK_CAMREFVALID : BOOL
VAR_INPUT
	CAMREF : MC_CAM_REF;
END_VAR
END_FUNCTION

(* ---- L_MB1P_CHECKREQUESTSINFO.pou ---- *)
FUNCTION L_MB1P_CHECKREQUESTSINFO : BOOL
VAR_OUTPUT
	XRTRIG : BOOL;
	XFTRIG : BOOL;
	DWRTRIG : DWORD;
	DWFTRIG : DWORD;
END_VAR
VAR_IN_OUT
	DWREQUESTSINFO : DWORD;
	DWREQUESTSINFO_OLD : DWORD;
END_VAR
END_FUNCTION

(* ---- L_MB1P_CONVERTDWORDTOLREALMODULOPOS.pou ---- *)
FUNCTION L_MB1P_CONVERTDWORDTOLREALMODULOPOS : LREAL
VAR_INPUT
	DWIN : DWORD;
	LRPERIOD : LREAL;
END_VAR
END_FUNCTION

(* ---- L_MB1P_CONVERTLREALTODWORDLMODULOPOS.pou ---- *)
FUNCTION L_MB1P_CONVERTLREALTODWORDLMODULOPOS : DWORD
VAR_INPUT
	LRIN : LREAL;
	LRPERIOD : LREAL;
END_VAR
END_FUNCTION

(* ---- L_MB1P_CONVERTPOSTOMODULOPOS.pou ---- *)
FUNCTION L_MB1P_CONVERTPOSTOMODULOPOS : LREAL
VAR_INPUT
	LRPOS : LREAL;
	LRPERIOD : LREAL;
END_VAR
VAR_OUTPUT
	DIREVCOUNTER : DINT;
END_VAR
END_FUNCTION

(* ---- L_MB1P_CONVERTPOSTOMODULOPOSEXTENDED.pou ---- *)
FUNCTION L_MB1P_CONVERTPOSTOMODULOPOSEXTENDED : LREAL
VAR_INPUT
	LRPOS : LREAL;
	LRPERIOD : LREAL;
END_VAR
VAR_OUTPUT
	DIREVCOUNTER : DINT;
END_VAR
END_FUNCTION

(* ---- L_MB1P_CONVERTPOSTOMODULOPOSFMOD.pou ---- *)
FUNCTION L_MB1P_CONVERTPOSTOMODULOPOSFMOD : LREAL
VAR_INPUT
	LRPOS : LREAL;
	LRPERIOD : LREAL;
END_VAR
END_FUNCTION

(* ---- L_MB1P_DIV.pou ---- *)
FUNCTION L_MB1P_DIV : LREAL
VAR_INPUT
	A : LREAL;
	B : LREAL;
END_VAR
END_FUNCTION

(* ---- L_MB1P_GETOVERRIDEFADINGTIME.pou ---- *)
FUNCTION L_MB1P_GETOVERRIDEFADINGTIME : BOOL
VAR_IN_OUT
	AXESGROUP : AXES_GROUP_KIN;
	WNUMOFMOVEFBS : WORD;
	LROVERRIDEFADINGTIME : LREAL;
	LRMAXVEL : LREAL := 0;
	LRMAXACC : LREAL := 0;
	LRMAXDEC : LREAL := 0;
	LRMAXJERK : LREAL := 0;
END_VAR
END_FUNCTION

(* ---- L_MB1P_GETPROFILETIMEMOVECONTPATH.pou ---- *)
FUNCTION L_MB1P_GETPROFILETIMEMOVECONTPATH : LREAL
VAR_IN_OUT
	AXESGROUP : AXES_GROUP_KIN;
	FB_MOVECONTPATH : L_MC4P_MoveContPath;
END_VAR
END_FUNCTION

(* ---- L_MB1P_GETTASKCYCLE.pou ---- *)
FUNCTION L_MB1P_GETTASKCYCLE : LREAL
END_FUNCTION

(* ---- L_MB1P_HLPCALCKOEFPOLY5THORD.pou ---- *)
FUNCTION L_MB1P_HLPCALCKOEFPOLY5THORD : ARRAY [0..5] OF LREAL
VAR_INPUT
	LRYPOSSTART : LREAL;
	LRYVELSTART : LREAL;
	LRYACCSTART : LREAL;
	LRYPOSEND : LREAL;
	LRYVELEND : LREAL;
	LRYACCEND : LREAL;
END_VAR
VAR_OUTPUT
	ALRKOEF : ARRAY [0..5] OF LREAL;
END_VAR
END_FUNCTION

(* ---- L_MB1P_HLPCALCYOFPOLY5THORDBASE.pou ---- *)
FUNCTION L_MB1P_HLPCALCYOFPOLY5THORDBASE : LREAL
VAR_OUTPUT
	LRYPOSSCALED : LREAL;
END_VAR
VAR_IN_OUT
	LRXPOSSCALED : LREAL;
	ALRKOEF : ARRAY [0..5] OF LREAL;
END_VAR
END_FUNCTION

(* ---- L_MB1P_HLPCALCYOFPOLY5THORDSTATE.pou ---- *)
FUNCTION L_MB1P_HLPCALCYOFPOLY5THORDSTATE : LREAL
VAR_INPUT
	LRXPOSSTART : LREAL;
	LRXPOSEND : LREAL := 1;
	LRSETXPOS : LREAL;
	ALRKOEF : ARRAY [0..5] OF LREAL;
END_VAR
VAR_OUTPUT
	LRYPOSSCALED : LREAL;
END_VAR
END_FUNCTION

(* ---- L_MB1P_HLPCHECKDIRECTION.pou ---- *)
FUNCTION L_MB1P_HLPCHECKDIRECTION : INT
VAR_IN_OUT
	LRPOSFIFOX : ARRAY [1..20] OF LREAL;
	LRLEN : LREAL;
END_VAR
END_FUNCTION

(* ---- L_MB1P_HLPDELTAVELTIMEEXTENDED.pou ---- *)
FUNCTION L_MB1P_HLPDELTAVELTIMEEXTENDED : BOOL
VAR_INPUT
	LRVELSTART : LREAL;
	LRACCSTART : LREAL;
	LRMAXACC : LREAL;
	LRMAXJERK : LREAL;
END_VAR
VAR_OUTPUT
	LRTIME : LREAL;
	LRDIST : LREAL;
END_VAR
END_FUNCTION

(* ---- L_MB1P_HLPDELTAVELTIMESTATE.pou ---- *)
FUNCTION L_MB1P_HLPDELTAVELTIMESTATE : BOOL
VAR_INPUT
	LRVELSTART : LREAL;
	LRACCSTART : LREAL;
	LRVELTARGET : LREAL;
	LRACCTARGET : LREAL;
	LRMAXACC : LREAL;
	LRMAXDEC : LREAL;
	LRMAXJERK : LREAL;
END_VAR
VAR_OUTPUT
	LRTIME : LREAL;
	LRDIST : LREAL;
END_VAR
END_FUNCTION

(* ---- L_MB1P_HLPDELTAVELTIMETOCONTANTVEL.pou ---- *)
FUNCTION L_MB1P_HLPDELTAVELTIMETOCONTANTVEL : BOOL
VAR_INPUT
	LRACCSTART : LREAL;
	LRMAXJERK : LREAL;
	WMODE : WORD;
END_VAR
VAR_OUTPUT
	LRVEL : LREAL;
	LRTIME : LREAL;
	LRDIST : LREAL;
END_VAR
END_FUNCTION

(* ---- L_MB1P_HLPDYNAMIZE.pou ---- *)
FUNCTION L_MB1P_HLPDYNAMIZE : LREAL
VAR_INPUT
	LRDIFF : LREAL;
	LRTIME : LREAL;
	LRCYCLETIME : LREAL;
END_VAR
END_FUNCTION

(* ---- L_MB1P_HLPFITCYCLE.pou ---- *)
FUNCTION L_MB1P_HLPFITCYCLE : LREAL
VAR_INPUT
	LRPOS : LREAL;
	LRLEN : LREAL;
END_VAR
END_FUNCTION

(* ---- L_MB1P_HLPFITCYCLELIM.pou ---- *)
FUNCTION L_MB1P_HLPFITCYCLELIM : BOOL
VAR_INPUT
	PLRPOS : POINTER TO LREAL;
	LRLEN : LREAL;
END_VAR
END_FUNCTION

(* ---- L_MB1P_HLPGEARRES.pou ---- *)
FUNCTION L_MB1P_HLPGEARRES : LREAL
VAR_INPUT
	LRINPUT : LREAL;
	LRNUM : LREAL;
	LRDEN : LREAL;
END_VAR
END_FUNCTION

(* ---- L_MB1P_HLPISLIMITED.pou ---- *)
FUNCTION L_MB1P_HLPISLIMITED : BOOL
VAR_INPUT
	LRVAL : LREAL;
END_VAR
END_FUNCTION

(* ---- L_MB1P_HLPMODULOADD.pou ---- *)
FUNCTION L_MB1P_HLPMODULOADD : LREAL
VAR_INPUT
	LRINPUT : LREAL;
	LROFFSET : LREAL;
	LRLENGHT : LREAL;
END_VAR
END_FUNCTION

(* ---- L_MB1P_HLPMODULODIFF.pou ---- *)
FUNCTION L_MB1P_HLPMODULODIFF : LREAL
VAR_INPUT
	LRDIFF : LREAL;
	LRLEN : LREAL;
END_VAR
END_FUNCTION

(* ---- L_MB1P_HLPMODULOOFFSET.pou ---- *)
FUNCTION L_MB1P_HLPMODULOOFFSET : LREAL
VAR_INPUT
	LROFFSET : LREAL;
	LRLENGTH : LREAL;
	PLROFFSETBASE : POINTER TO LREAL;
END_VAR
END_FUNCTION

(* ---- L_MB1P_HLPMODULOSUB.pou ---- *)
FUNCTION L_MB1P_HLPMODULOSUB : LREAL
VAR_INPUT
	LRDIFF : LREAL;
	LRLEN : LREAL;
END_VAR
END_FUNCTION

(* ---- L_MB1P_HLPMODULOZEROPOS.pou ---- *)
FUNCTION L_MB1P_HLPMODULOZEROPOS : BOOL
VAR_INPUT
	PLRPOS : POINTER TO LREAL;
	LRLENINT : LREAL;
END_VAR
END_FUNCTION

(* ---- L_MB1P_HLPPOLY4RG.pou ---- *)
FUNCTION L_MB1P_HLPPOLY4RG : LREAL
VAR_INPUT
	LRX : LREAL;
END_VAR
END_FUNCTION

(* ---- L_MB1P_HLPPT1FILT.pou ---- *)
FUNCTION L_MB1P_HLPPT1FILT : LREAL
VAR_INPUT
	LRVALUE : LREAL;
	LRINPUT : LREAL;
	LRNEW_N : LREAL;
END_VAR
END_FUNCTION

(* ---- L_MB1P_HLPSIGNNE.pou ---- *)
FUNCTION L_MB1P_HLPSIGNNE : BOOL
VAR_INPUT
	A : LREAL;
	B : LREAL;
END_VAR
END_FUNCTION

(* ---- L_MB1P_IDENTMAXPOSSIBLEDIAMETER.pou ---- *)
FUNCTION L_MB1P_IDENTMAXPOSSIBLEDIAMETER : LREAL
VAR_INPUT
	WIDENTDIAMCALCCYCLES : WORD := 1;
END_VAR
VAR_IN_OUT
	LRACTDANCERPOSIN : LREAL;
	LRMAXDANCERPOS : LREAL;
	LRDANCERMATERIALLENGTH : LREAL;
	LRDIAMCALCDIST : LREAL;
END_VAR
END_FUNCTION

(* ---- L_MB1P_LREQ.pou ---- *)
FUNCTION L_MB1P_LREQ : BOOL
VAR_INPUT
	LRVALUE : LREAL;
	LRTARGET : LREAL;
END_VAR
END_FUNCTION

(* ---- L_MB1P_LRGE.pou ---- *)
FUNCTION L_MB1P_LRGE : BOOL
VAR_INPUT
	LRVALUE : LREAL;
	LRTARGET : LREAL;
END_VAR
END_FUNCTION

(* ---- L_MB1P_LRGT.pou ---- *)
FUNCTION L_MB1P_LRGT : BOOL
VAR_INPUT
	LRVALUE : LREAL;
	LRTARGET : LREAL;
END_VAR
END_FUNCTION

(* ---- L_MB1P_LRLE.pou ---- *)
FUNCTION L_MB1P_LRLE : BOOL
VAR_INPUT
	LRVALUE : LREAL;
	LRTARGET : LREAL;
END_VAR
END_FUNCTION

(* ---- L_MB1P_LRLT.pou ---- *)
FUNCTION L_MB1P_LRLT : BOOL
VAR_INPUT
	LRVALUE : LREAL;
	LRTARGET : LREAL;
END_VAR
END_FUNCTION

(* ---- L_MB1P_LRNE.pou ---- *)
FUNCTION L_MB1P_LRNE : BOOL
VAR_INPUT
	LRVALUE : LREAL;
	LRTARGET : LREAL;
END_VAR
END_FUNCTION

(* ---- L_MB1P_MODULOCYCLE.pou ---- *)
FUNCTION L_MB1P_MODULOCYCLE : LREAL
VAR_INPUT
	LRPOSIN : LREAL;
	LRPOSITIONPERIOD : LREAL;
END_VAR
END_FUNCTION

(* ---- L_MB1P_POSITIONINSIDEWINDOW.pou ---- *)
FUNCTION L_MB1P_POSITIONINSIDEWINDOW : BOOL
VAR_INPUT
	LRPOSIN : LREAL;
	LRLOWERWINDOW : LREAL;
	LRUPPERWINDOW : LREAL;
END_VAR
VAR_OUTPUT
	XERROR : BOOL := FALSE;
END_VAR
VAR_IN_OUT
	AXIS : AXIS_REF;
END_VAR
END_FUNCTION

(* ---- L_MB1P_PROFILETIMEVALID.pou ---- *)
FUNCTION L_MB1P_PROFILETIMEVALID : BOOL
VAR_IN_OUT
	LRPROFILETIME : LREAL;
END_VAR
END_FUNCTION

(* ---- L_TT1P_CALCSYNCTIME.pou ---- *)
FUNCTION L_TT1P_CALCSYNCTIME : BOOL
VAR_INPUT
	LRACTMATERIALVEL : LREAL;
	LRACCMAX : LREAL;
	LRJERKSTART : LREAL;
	LRJERKEND : LREAL;
END_VAR
VAR_OUTPUT
	LRACCTIME : LREAL;
	LRACCDIST : LREAL;
END_VAR
END_FUNCTION

(* ---- SB_CALCULATEPRODUCTERROR.pou ---- *)
FUNCTION SB_CALCULATEPRODUCTERROR : LREAL
VAR_INPUT
	LRPRODUCTTARGETCORRECTED : LREAL;
	LRMASTERPOSITIONATDETECTION : LREAL;
	LRCORRECTEDFACTORCOMPAREPOSITION : LREAL;
	BYNUMBEROFTARGETS : BYTE;
	LRMASTERCYCLELENGTH : LREAL;
END_VAR
END_FUNCTION

(* ---- _L_MB1A_ANALOGINTOSPEEDOUT.pou ---- *)
FUNCTION_BLOCK _L_MB1A_ANALOGINTOSPEEDOUT
VAR_INPUT
	WINPUT : WORD;
	WUPPERLIM : WORD := 16000;
	WLOWERLIM : WORD := 0;
	LRUPPERSPEEDLIM : LREAL := 1000.0;
	LRLOWERSPEEDLIM : LREAL := -1000.0;
	RFILTTIME : REAL := 0.01;
	LRACC : LREAL := 1000;
	LRDEC : LREAL := 1000;
	LRJERK : LREAL := 100000;
	XNEGATIVEDIRECTION : BOOL;
	LRDEADBANDWINDOW : LREAL := 10;
END_VAR
VAR_OUTPUT
	LRSETSPEEDOUT : LREAL;
END_VAR
VAR
	LRSPEEDSETPOINT : LREAL;
	L_MB1P_RAMPGENERATOR1 : L_MC1P_RampGenerator;
END_VAR
END_FUNCTION_BLOCK

(* ---- _L_MB1A_IOSELECTMASK.pou ---- *)
FUNCTION_BLOCK _L_MB1A_IOSELECTMASK
VAR_INPUT
	XENABLE : BOOL;
	WNUMOFMASK : WORD := 3;
	XSELECTMASK : BOOL;
	XIP1 : BOOL;
	XIP2 : BOOL;
	XIP3 : BOOL;
	XIP4 : BOOL;
	XIP5 : BOOL;
	XIP6 : BOOL;
	XIP7 : BOOL;
	XIP8 : BOOL;
END_VAR
VAR_OUTPUT
	XBLINKEROUT : BOOL;
	WNOOUT : WORD;
	WMASK : WORD;
	AXOP1 : ARRAY [1..10] OF BOOL;
	AXOP2 : ARRAY [1..10] OF BOOL;
	AXOP3 : ARRAY [1..10] OF BOOL;
	AXOP4 : ARRAY [1..10] OF BOOL;
	AXOP5 : ARRAY [1..10] OF BOOL;
	AXOP6 : ARRAY [1..10] OF BOOL;
	AXOP7 : ARRAY [1..10] OF BOOL;
	AXOP8 : ARRAY [1..10] OF BOOL;
END_VAR
VAR
	XSELECTMASK_OLD : BOOL;
	XBLINKEROUT_OLD : BOOL;
	TON_1 : TON;
	TOF_1 : TOF := STRUCT(PT := TIME#400ms);
	WCNTR : WORD;
	XBLINKER : BOOL;
	XIP1_OLD : BOOL;
	XIP2_OLD : BOOL;
	XIP3_OLD : BOOL;
	XIP4_OLD : BOOL;
	XIP5_OLD : BOOL;
	XIP6_OLD : BOOL;
	XIP7_OLD : BOOL;
	XIP8_OLD : BOOL;
END_VAR
END_FUNCTION_BLOCK

METHOD CALL_BLINKER
END_METHOD

(* ---- _L_MB1P_ANALOGINPUTSPEEDCTRL.pou ---- *)
FUNCTION_BLOCK _L_MB1P_ANALOGINPUTSPEEDCTRL
VAR_INPUT
	WINPUT : WORD;
	WUPPERLIM : WORD := 10000;
	WLOWERLIM : WORD := 0;
	LRUPPERSPEEDLIM : LREAL := 1000;
	LRLOWERSPEEDLIM : LREAL := 0;
	LRDEADBAND : LREAL := 5;
	RFILTTIME : REAL := 0.01;
	LRACC : LREAL := 1000;
	LRDEC : LREAL := 1000;
	LRJERK : LREAL := 100000;
	XNEGATIVEDIRECTION : BOOL;
END_VAR
VAR_OUTPUT
	LRSETSPEEDOUT : LREAL;
END_VAR
VAR
	LRINPUTSCALED : LREAL;
	LRSPEEDSETPOINT : LREAL;
	L_D94A_FILTER : L_USPP_PT1Filter;
	L_MB1P_RAMPGENERATOR1 : L_MC1P_RampGenerator;
END_VAR
END_FUNCTION_BLOCK

(* ---- _L_MB1P_AXISCONTROLBYPOS.pou ---- *)
FUNCTION_BLOCK _L_MB1P_AXISCONTROLBYPOS
VAR_INPUT
	XENABLE : BOOL;
	LRSETPOSITION : LREAL;
	LRSETVELOCITY : LREAL;
	LRSETACCELERATION : LREAL;
	ESETVALUEMODE : L_MC1P_SetValueMode := L_MC1P_SetValueMode.Pos;
END_VAR
VAR_OUTPUT
	XBUSY : BOOL;
	XCOMMANDABORTED : BOOL;
	XERROR : BOOL;
	EERRORID : L_IE1P_Error;
	LRSETPOSOUT : LREAL;
END_VAR
VAR_IN_OUT
	AXIS : AXIS_REF;
END_VAR
VAR
	LRSETPOSITION_INT : LREAL;
	XENABLE_OLD : BOOL;
	XBUSY_OLD : BOOL;
	ESTATE : L_MB1P_States;
	MC_HALT1 : MC_HALT;
	FB_FOLLOWSETVALUES : L_MC1P_FollowSetValues;
END_VAR
END_FUNCTION_BLOCK

METHOD CALL_ERRORHANDLER
END_METHOD

METHOD CALL_FBMETHODS
END_METHOD

METHOD CALL_FB_FOLLOWSETVALUES
END_METHOD

METHOD CALL_MC_HALT
END_METHOD

METHOD CALL_MC_HALT_INPUT
END_METHOD

METHOD CALL_OUTPUT
END_METHOD

METHOD CALL_RESETCOMMANDS
END_METHOD

METHOD CALL_RESETOUTPUT
END_METHOD

METHOD CALL_STATEMACHINE
END_METHOD

METHOD CALL_S000_CYCLIC
END_METHOD

METHOD CALL_S001_INIT
END_METHOD

METHOD CALL_S002_READY
END_METHOD

METHOD CALL_S999_ERROR
END_METHOD

(* ---- _L_MB1P_AXISCONTROLBYVEL.pou ---- *)
FUNCTION_BLOCK _L_MB1P_AXISCONTROLBYVEL
VAR_INPUT
	XENABLE : BOOL;
	LRSETVELOCITY : LREAL;
END_VAR
VAR_OUTPUT
	XBUSY : BOOL;
	XCOMMANDABORTED : BOOL;
	XERROR : BOOL;
	EERRORID : L_IE1P_Error;
	LRSETVELOUT : LREAL;
END_VAR
VAR_IN_OUT
	AXIS : AXIS_REF;
END_VAR
VAR
	LRSETVELOCITY_INT : LREAL;
	XENABLE_OLD : BOOL;
	XBUSY_OLD : BOOL;
	ESTATE : L_MB1P_States;
	MC_HALT1 : MC_HALT;
	FB_FOLLOWSETVALUES : L_MC1P_FollowSetValues;
END_VAR
END_FUNCTION_BLOCK

METHOD CALL_ERRORHANDLER
END_METHOD

METHOD CALL_FBMETHODS
END_METHOD

METHOD CALL_FB_FOLLOWSETVALUES
END_METHOD

METHOD CALL_MC_HALT
END_METHOD

METHOD CALL_MC_HALT_INPUT
END_METHOD

METHOD CALL_OUTPUT
END_METHOD

METHOD CALL_RESETCOMMANDS
END_METHOD

METHOD CALL_RESETOUTPUT
END_METHOD

METHOD CALL_STATEMACHINE
END_METHOD

METHOD CALL_S000_CYCLIC
END_METHOD

METHOD CALL_S001_INIT
END_METHOD

METHOD CALL_S002_READY
END_METHOD

METHOD CALL_S999_ERROR
END_METHOD
